(* IEC 61131-3 sources: daoli-st-library/DL_Base (part 14) *)

(* ---- FB_DL_MutexOwnerAudit.st ---- *)
(*
  FB_DL_MutexOwnerAudit  —  互斥锁所有权审计台账 / Mutex ownership audit ledger
  分类 Category : DL_Base
  码位 Code     : 16#01_0_02
  段位说明      : 01_0 段仅占 00/01（R38），02 起空穴，本件启用 02 格
  版本 Version  : 1.0.1
  来源 Source   : t0-8-sema — T0-8 行待挖子项「超时归还后的所有权审计」落地
  溯源 Origin   : clean-room 实现，未复制任何源码行
  功能 Function : 1) 只做「事后可追」审计出口，不改变加解锁语义：与 FB_DL_SemaMutex（互斥本体）
                  分工，本体管仲裁，本件管台账；
                  2) 记录持锁者标识 uOwnerCur、当前持有时长 fHoldCurSec、累计持有时长 uHoldTotalSec；
                  3) 计数台账：申请 / 正常释放 / 越权释放 / 超时强制归还四类，全部饱和计数不回绕；
                  4) 越权释放（无主时的释放沿）记故障级码并锁存，bReset 解除；
                  5) 超时强制归还由调用方把 FB_DL_SemaMutex.bTimedOut 单拍脉冲接入 bTimeoutForced。
  边界 Boundary : ① 本件不仲裁、不拒绝任何事件，只记录；仲裁语义全部由 FB_DL_SemaMutex 承载；
                  ② uDeltaTimeMs 为调用方注入的任务周期 [ms]，越界按上限钳位（防一次错误注入污染台账）；
                  R41 返修（R241）：饱和闸整体上移 UDINT 域——加法前预留量预检
                  （_uHoldMs / _uHoldTotMs 各自与 DL_MUA_MS_MAX - _uDtEff 比较），
                  判定值域 0..16#FFFF_F000 ms（约 49.7 天），以 10 ms 任务周期计约
                  4.29 亿拍可达，饱和分支真实可达，秒换算改纯 UDINT 整除，零降型路径；
                  ③ uOwnerIdClaim = 0 视为非法标识：照常记录持有但置信息级码 0302；
                  ④ 审计状态两相 CASE 全覆盖 + ELSE 兜底；无定时器/边沿以外的时序假设。
  依赖 Depends  : 仅 Standard.library（R_TRIG）；与 FB_DL_SemaMutex（已注册）仅状态语义对齐，不实例化
  码表 Error codes（本件格 01_0_02，子码步进 +0x100）:
    16#0001_0102 信息级：本拍记录到申请沿（持锁开始）
    16#0001_0202 故障级：越权释放（无主时的释放沿），锁存至 bReset
    16#0001_0302 信息级：申请者标识非法（uOwnerIdClaim = 0），记录照常完成
    16#0001_0402 信息级：超时强制归还事件已入账
    16#0001_0502 故障级：审计相位落 ELSE 兜底（非法相位 ID），强制回无主相并锁存

  修订历史 Revision :
    2026-11-19  v1.0.0  R39 首版（批次 1 · 序号 1）
    2026-11-19  v1.0.1  R40 5 抽终审挂账（不改逻辑）：⚠ 段 4 行 108 饱和闸「UDINT_TO_DINT(DL_MUA_SEC_MAX)」
                  对 16#FFFF_FFFE 做 DINT 降型溢出（回绕为负），乘积类型跨平台歧义；且 _uHoldTotMs
                  （UDINT ms）数学上不可能达到 SEC_MAX×1000 ms，秒级饱和分支永不按预期触发，返修轮处理。
    2026-11-19  v1.0.1  R41 P0-2 返修实施：删除「UDINT_TO_DINT(SEC_MAX) × 1000」降型比较与
                  不可达秒级闸，改为 UDINT 域加法前预留量预检（判定值域 0..16#FFFF_F000 ms，
                  可达性向量已写入边界②），秒换算改纯 UDINT 整除；新增常量 DL_MUA_MS_MAX，
                  DL_MUA_SEC_MAX 降级为文档口径不再参与比较。
*)

TYPE E_DL_MutexAuditState :
(
    eFree := 0,    // 无主：互斥空闲，等待申请沿 / Free, mutex idle, waiting for a claim edge
    eHeld := 10    // 有主：持锁审计中，累计持有时长 / Held, ownership held and hold time accumulating
);
END_TYPE

FUNCTION_BLOCK FB_DL_MutexOwnerAudit
VAR_INPUT
    bClaimEvt      : BOOL;                  // 申请事件沿（来自本体申请沿或其输入 CLK）[-] / Claim event edge from the mutex body
    bReleaseEvt    : BOOL;                  // 释放事件沿（来自本体释放沿或其输入 CLK）[-] / Release event edge from the mutex body
    bTimeoutForced : BOOL;                  // 超时强制归还脉冲，接 FB_DL_SemaMutex.bTimedOut 单拍输出 [-] / Forced timeout return pulse, wire SemaMutex.bTimedOut
    uOwnerIdClaim  : DINT := 0;             // 本次申请者标识 [ID]，0 = 非法（置信息码） / Claimer owner ID, 0 = illegal (info code)
    uDeltaTimeMs   : UDINT := 10;           // 任务周期注入 [ms]，越界按上限钳位 / Task cycle time injected by caller [ms]
    bReset         : BOOL := FALSE;         // 审计复位，上升沿清越权锁存（不清台账计数）/ Audit reset, rising edge clears the fault latch only
END_VAR
VAR_OUTPUT
    eState         : E_DL_MutexAuditState;  // 审计状态出口，段尾单点映射 / Audit state outlet
    bHeld          : BOOL;                  // 当前有主（与 eHeld 同源派生）/ Mutex currently held, derived from eHeld
    uOwnerCur      : DINT;                  // 当前持锁者标识 [ID]，无主时为 0 / Current owner ID, 0 when free
    fHoldCurSec    : REAL;                  // 当前连续持有时长 [s]，释放拍冻结到释放值 / Current continuous hold time [s], frozen at release
    uHoldTotalSec  : UDINT;                 // 累计持有时长 [s]，饱和不回绕 / Total accumulated hold time [s], saturating
    uClaimCnt      : UDINT;                 // 累计申请次数 [次]，饱和不回绕 / Total claim count [times], saturating
    uReleaseCnt    : UDINT;                 // 累计正常释放次数 [次]，饱和不回绕 / Total normal release count [times], saturating
    uUnauthRelCnt  : UDINT;                 // 累计越权释放次数 [次]，饱和不回绕 / Total unauthorized release count [times], saturating
    uTimeoutCnt    : UDINT;                 // 累计超时强制归还次数 [次]，饱和不回绕 / Total forced timeout return count [times], saturating
    uErrorId       : UDINT;                 // 事件码，0 = 无事件（故障级码锁存回放）/ Event code, 0 = none, fault codes latched and replayed
END_VAR
VAR
    rtClaim        : R_TRIG;                // 申请沿实例，主体首部无条件刷新 / Claim edge instance, refreshed unconditionally
    rtRelease      : R_TRIG;                // 释放沿实例，主体首部无条件刷新 / Release edge instance, refreshed unconditionally
    rtTimeout      : R_TRIG;                // 超时归还沿实例，主体首部无条件刷新 / Timeout edge instance, refreshed unconditionally
    rtReset        : R_TRIG;                // 复位沿实例，主体首部无条件刷新 / Reset edge instance, refreshed unconditionally
    _eState        : E_DL_MutexAuditState := E_DL_MutexAuditState.eFree;  // 内部审计相位（CASE 唯一写入目标）/ Internal audit phase, sole CASE target
    _uFault        : UDINT;                 // 故障码锁存寄存 / Latched fault code register
    _uInfo         : UDINT;                 // 本拍信息码，每拍重算 / Transient info code this cycle
    _uOwnerInt     : DINT := 0;             // 内部持锁者标识，对外经 uOwnerCur 镜像 / Internal owner register mirrored to uOwnerCur
    _uHoldMs       : UDINT := 0;            // 当前持有毫秒累加器 [ms] / Current hold millisecond accumulator
    _uHoldTotMs    : UDINT := 0;            // 累计持有毫秒累加器 [ms] / Total hold millisecond accumulator
    _uDtEff        : UDINT;                 // 钳位后的生效周期 [ms] / Clamped effective cycle time
END_VAR
VAR CONSTANT
    DL_MUA_DT_MAX     : UDINT := 60000;         // 单拍周期合理上限 [ms]，超出按上限入账 / Sane per-cycle cap [ms]
    DL_MUA_CNT_MAX    : UDINT := 16#FFFF_FFFE;  // 各计数饱和上限 [次]，加一永不回绕 / Counter saturation bound, increment never wraps
    DL_MUA_MS_PER_SEC : UDINT := 1000;          // 每秒毫秒数 [ms/s] / Milliseconds per second
    DL_MUA_SEC_MAX    : UDINT := 16#FFFF_FFFE;  // 秒级累计饱和上限 [s]，R41 起仅作文档口径，不再参与比较 / Second-level doc bound, not used in comparison since R41
    DL_MUA_MS_MAX     : UDINT := 16#FFFF_F000;  // 毫秒累加器饱和上限 [ms]，UDINT 域加法闸（约 49.7 天，10ms 周期约 4.29 亿拍可达）/ Millisecond accumulator saturation bound, UDINT-domain add gate
END_VAR

(* —— 段 0：边沿实例无条件周期刷新（R7 红线：严禁置于 IF/CASE 分支内） —— *)
rtClaim(CLK := bClaimEvt);                                        // 申请沿刷新，每拍必调
rtRelease(CLK := bReleaseEvt);                                    // 释放沿刷新，每拍必调
rtTimeout(CLK := bTimeoutForced);                                 // 超时归还沿刷新，每拍必调
rtReset(CLK := bReset);                                           // 复位沿刷新，每拍必调

(* —— 段 1：单拍量预清零（锁存量 _uFault 与台账计数不入清单，R187①） —— *)
_uInfo := 16#0000_0000;             // 信息码每拍重算
_uFault := _uFault;                 // 故障锁存码保持回放（禁同拍抹除，R187/R189）
uErrorId := 16#0000_0000;           // 事件码缺省无事件（段尾按锁存/信息单点回放）

(* —— 段 2：周期注入钳位（防御：一次错误注入不得污染台账） —— *)
IF uDeltaTimeMs > DL_MUA_DT_MAX THEN
    _uDtEff := DL_MUA_DT_MAX;       // 越界按上限钳位
ELSE
    _uDtEff := uDeltaTimeMs;        // 域内直通
END_IF

(* —— 段 3：复位沿（只清越权锁存，不清台账计数——台账是历史事实） —— *)
IF rtReset.Q THEN
    _uFault := 16#0000_0000;        // 清故障锁存码（唯一解除路径：bReset 上升沿）
END_IF

(* —— 段 4：持有时长累加（仅 eHeld 相累计；R41 P0-2 返修：饱和闸整体上移 UDINT 域，
     加法前预留量预检，判定值域 0..16#FFFF_F000 ms，无降型、无可达性缺口） —— *)
IF _eState = E_DL_MutexAuditState.eHeld THEN
    IF _uHoldMs <= DL_MUA_MS_MAX - _uDtEff THEN     // 加前预留量预检（当拍量判据，UDINT 域）
        _uHoldMs := _uHoldMs + _uDtEff;             // 当前持有累加 [ms]
    ELSE
        _uHoldMs := DL_MUA_MS_MAX;                  // 饱和钳位，永不回绕
    END_IF
    IF _uHoldTotMs <= DL_MUA_MS_MAX - _uDtEff THEN  // 同口径预检累计累加器（UDINT 域，零降型）
        _uHoldTotMs := _uHoldTotMs + _uDtEff;       // 累计持有累加 [ms]
    ELSE
        _uHoldTotMs := DL_MUA_MS_MAX;               // 累计饱和钳位，永不回绕
    END_IF
END_IF
fHoldCurSec := UDINT_TO_REAL(_uHoldMs) / UDINT_TO_REAL(DL_MUA_MS_PER_SEC);  // 当前持有换算秒（分母为常量恒非零）
uHoldTotalSec := _uHoldTotMs / DL_MUA_MS_PER_SEC;   // 累计秒整除换算（纯 UDINT 域，R241 零降型）

(* —— 段 5：审计相位机（只记录、不仲裁；出口在段 7） —— *)
CASE _eState OF

E_DL_MutexAuditState.eFree:
    IF rtRelease.Q THEN
        uUnauthRelCnt := uUnauthRelCnt + 1;     // 越权释放入账（无主时的释放沿）
        IF uUnauthRelCnt >= DL_MUA_CNT_MAX THEN
            uUnauthRelCnt := DL_MUA_CNT_MAX;    // 计数饱和防回绕
        END_IF
        _uFault := 16#0001_0202;                // 故障级：越权释放，锁存至 bReset
    ELSIF rtTimeout.Q THEN
        uTimeoutCnt := uTimeoutCnt + 1;         // 超时归还沿落在此相同样入账（本体已强制归还）
        IF uTimeoutCnt >= DL_MUA_CNT_MAX THEN
            uTimeoutCnt := DL_MUA_CNT_MAX;
        END_IF
        _uInfo := 16#0001_0402;                 // 信息级：超时归还已入账
    ELSIF rtClaim.Q THEN
        uClaimCnt := uClaimCnt + 1;             // 申请入账
        IF uClaimCnt >= DL_MUA_CNT_MAX THEN
            uClaimCnt := DL_MUA_CNT_MAX;
        END_IF
        IF uOwnerIdClaim = 0 THEN
            _uInfo := 16#0001_0302;             // 信息级：标识非法，记录照常
        ELSE
            _uInfo := 16#0001_0102;             // 信息级：持锁开始
        END_IF
        _uOwnerInt := uOwnerIdClaim;            // 记录持锁者标识（含非法 0，照实记录）
        _uHoldMs := 0;                          // 当前持有时长从零起算
        _eState := E_DL_MutexAuditState.eHeld;  // 进有主相
    END_IF

E_DL_MutexAuditState.eHeld:
    IF rtRelease.Q THEN
        uReleaseCnt := uReleaseCnt + 1;         // 正常释放入账
        IF uReleaseCnt >= DL_MUA_CNT_MAX THEN
            uReleaseCnt := DL_MUA_CNT_MAX;
        END_IF
        _uOwnerInt := 0;                        // 无主：标识清零
        _eState := E_DL_MutexAuditState.eFree;  // 回无主相（当前持有时长冻结在释放值）
    ELSIF rtTimeout.Q THEN
        uTimeoutCnt := uTimeoutCnt + 1;         // 超时强制归还有主相入账
        IF uTimeoutCnt >= DL_MUA_CNT_MAX THEN
            uTimeoutCnt := DL_MUA_CNT_MAX;
        END_IF
        _uInfo := 16#0001_0402;                 // 信息级：超时归还已入账
        _uOwnerInt := 0;                        // 强制归还：标识清零
        _eState := E_DL_MutexAuditState.eFree;  // 回无主相
    ELSIF rtClaim.Q THEN
        uClaimCnt := uClaimCnt + 1;             // 有主期间的申请沿照常入账（本体仲裁语义不变）
        IF uClaimCnt >= DL_MUA_CNT_MAX THEN
            uClaimCnt := DL_MUA_CNT_MAX;
        END_IF
    END_IF

ELSE
    _uFault := 16#0001_0502;                    // 故障级：非法相位 ID 兜底，锁存至 bReset
    _uOwnerInt := 0;                            // 无主侧强制清标识（安全侧）
    _eState := E_DL_MutexAuditState.eFree;      // 强制回无主相（自恢复，不锁死）

END_CASE

(* —— 段 6：派生输出每拍重写（名实同源） —— *)
bHeld := (_eState = E_DL_MutexAuditState.eHeld);            // 有主派生位
uOwnerCur := _uOwnerInt;                                     // 持锁者镜像输出

(* —— 段 7：事件码单点回放（故障锁存优先，信息码其次） —— *)
IF _uFault <> 16#0000_0000 THEN
    uErrorId := _uFault;            // 故障锁存码回放（不在故障态按当下输入重推）
ELSE
    uErrorId := _uInfo;             // 信息码
END_IF
eState := _eState;                  // 状态出口单点映射

END_FUNCTION_BLOCK

(* ---- FB_DL_OutputForcingBank.st ---- *)
(*==============================================================================
 * 组件名称 (Component)  : FB_DL_OutputForcingBank
 * 所属子库 (Sublibrary) : DL_Base
 * 当前版本 (Version)    : 1.0.0
 * 兼容性   (Platform)   : CODESYS 3.5+ / TwinCAT 3 / 汇川 InoProShop / 施耐德 Machine Expert
 *                         仅依赖 Standard.library（R_TRIG），零厂商私有库
 * 功能描述 (Function)   : 16 路输出强制库（调试/维修用）：每拍组合式裁决
 *                         abOut[i] = bAutoMode ∧ abForceSel[i] ? abForceVal[i]
 *                         : abAutoVal[i]；任一通道强制激活 → uForcingMask 位图
 *                         对应位置 1；强制撤除（abForceSel 下降沿）当拍无扰
 *                         回自动（组合式单拍重算，无斜坡无残留）；bAutoMode=
 *                         FALSE 时强制请求被拒（输出仍走自动值），拒收当拍置
 *                         信息码 eForceRej 并计数 uRejCnt。
 * 接口     (Interface)  : 输入 abAutoVal 16 路自动值、abForceSel 16 路强制选择、
 *                         abForceVal 16 路强制值、bAutoMode 自动模式许可；
 *                         输出 abOut 16 路裁决输出、uForcingMask 强制激活
 *                         位图（bit i=通道 i）、uRejCnt 强制拒收计数、
 *                         eErrCode 信息码、bError 故障标志（本件无故障级
 *                         条件，恒 FALSE，契约位保留）。
 * 边界     (Boundary)   : ① **属主边界（写死）：本件只做输出裁决，不接管安全
 *                         回路、不做强制权限管理**；安全回路强制归硬件层，
 *                         本件不得用于旁路安全联锁（头注释声明）。
 *                         ② 无扰回自动：撤除拍输出 = 自动值（组合式当拍生效，
 *                         无历史残留路径，规格指定）。
 *                         ③ 拒收计数用 R_TRIG 捕「拒收状态进入沿」计数（状态
 *                         电平不重复计数）；拒收期 uForcingMask 对应位保持 0
 *                         （强制未生效）。
 *                         ④ 通道定长 16（常量），FOR 界宽常量，无越界路径。
 *                         ⑤ R_TRIG 实例段 0 无条件周期调用（R6/R7）。
 *                         ⑥ 零全局耦合（无 GVL / VAR_EXTERNAL / 物理地址）。
 * 分工声明 (Scope)      : 与 `FB_DL_OverrideSelector` 分工：模拟量超驰选择归
 *                         那件、数字量强制库归本件；与 `FB_DL_InterlockMatrix`
 *                         分工：联锁矩阵归那件（安全语义），本件为非安全
 *                         调试设施。
 * 来源标签 (Source Tag) : 自研线（输出强制裁决为道莅防御性实现）
 * 码表     (Codes)      : 本件不占用任何全局数字码位。出口为 BOOL 数组 +
 *                         WORD 位图 + UDINT 计数 + ENUM 信息码；数字码位待
 *                         主控收口阶段统一派号。
 * 红线自检 (Redline)    : R1 ✓ 零 GVL/VAR_EXTERNAL ｜ R2 ✓ 零 %I/%Q/%M ｜ R3 ✓ 纯 IEC 61131-3
 *                         R4 ✓ 拒收沿计数 + 无扰回自动 + 位图单源 ｜ R5 ✓ 声明逐行同行双语注释
 *                         R6 N/A（无 ENUM 状态机） ｜ R7 ✓ 一 R_TRIG 段 0 无条件刷新
 * 修订历史 (Revision)   : 2026-11-20  v1.0.0  R50 首版（批次 3 · 序号 12）
 * 验收向量 (Acceptance) : ① bAutoMode=TRUE，abForceSel[3]=TRUE，abForceVal[3]=
 *                         TRUE，abAutoVal[3]=FALSE → abOut[3]=TRUE，
 *                         uForcingMask.bit3=1；② abForceSel[3] 撤除当拍：
 *                         abOut[3]=abAutoVal[3]=FALSE（无扰回自动），bit3=0；
 *                         ③ bAutoMode=FALSE 且 abForceSel[5] 置位 → abOut[5]
 *                         =abAutoVal[5]（强制被拒），uRejCnt+1，
 *                         eErrCode=eForceRej。
 *==============================================================================*)

(*-----------------------------------------------------------------------------
 * 枚举: E_DL_OfbErr（信息码；拒收走信息级，不置 bError）
 *----------------------------------------------------------------------------*)
TYPE E_DL_OfbErr :
(
    eOk       := 0,   // 无拒收 / No rejection
    eForceRej := 1    // 信息级：存在被拒强制通道（bAutoMode=FALSE，见 uRejCnt） / Info: forced channels rejected
);
END_TYPE

FUNCTION_BLOCK FB_DL_OutputForcingBank
VAR_INPUT
    abAutoVal  : ARRAY[0..15] OF BOOL;   // 16 路自动值（正常输出源） [-] / Sixteen auto values
    abForceSel : ARRAY[0..15] OF BOOL;   // 16 路强制选择 [-] / Sixteen force selects
    abForceVal : ARRAY[0..15] OF BOOL;   // 16 路强制值 [-] / Sixteen force values
    bAutoMode  : BOOL := TRUE;           // 自动模式许可（FALSE=强制被拒） [-] / Auto-mode permission
END_VAR
VAR_OUTPUT
    abOut        : ARRAY[0..15] OF BOOL; // 16 路裁决输出 [-] / Sixteen arbitrated outputs
    uForcingMask : WORD;                 // 强制激活位图（bit i=通道 i 强制生效） [-] / Forcing bitmap
    uRejCnt      : UDINT := 0;           // 强制拒收进入沿计数（防回绕） [次] / Rejection entry count
    eErrCode     : E_DL_OfbErr;          // 信息码出口 / Info code outlet
    bError       : BOOL;                 // 故障标志（本件恒 FALSE，契约位） [-] / Error flag, contract pin, always FALSE
END_VAR
VAR
    _uMask    : WORD;                    // 位图内部单源（与出口同源） / Bitmap internal source
    _bAnyRej  : BOOL;                    // 存在拒收通道当拍量 [-] / Any rejected channel
    i         : DINT;                    // 通道循环索引 / Channel loop index
    rtRej     : R_TRIG;                  // 拒收进入沿实例，段 0 无条件调用 / Rejection entry edge instance
END_VAR
VAR CONSTANT
    DL_OFB_NMAX : DINT := 16;            // 通道定长 [路] / Fixed channel count
    DL_OFB_BIT0 : WORD := 1;             // bit0 基准掩码 [-] / Bit zero base mask
    DL_OFB_UDMAX: UDINT := 4294967295;   // 拒收计数饱和点（防回绕） [次] / Rejection counter ceiling
END_VAR

(* —— 段 0：拒收沿实例无条件周期刷新（R6/R7） —— *)
rtRej(CLK := (NOT bAutoMode) AND (abForceSel[0] OR abForceSel[1] OR abForceSel[2]
       OR abForceSel[3] OR abForceSel[4] OR abForceSel[5] OR abForceSel[6]
       OR abForceSel[7] OR abForceSel[8] OR abForceSel[9] OR abForceSel[10]
       OR abForceSel[11] OR abForceSel[12] OR abForceSel[13] OR abForceSel[14]
       OR abForceSel[15]));              // 拒收进入沿（任一强制选择 ∧ 非自动模式），每拍必调 / Rejection entry edge, every scan

(* —— 段 1：拒收沿计数（防回绕） —— *)
IF rtRej.Q THEN
    IF uRejCnt < DL_OFB_UDMAX THEN
        uRejCnt := uRejCnt + 1;          // 拒收进入沿计数 / Count rejection entry
    END_IF
END_IF

(* —— 段 2：16 路组合式裁决（强制生效闸：bAutoMode ∧ abForceSel；撤除当拍无扰回自动） —— *)
_uMask := 0;                             // 位图当拍重建（单源） / Rebuild bitmap per scan
_bAnyRej := FALSE;                       // 拒收量预清 / Rejection preset
FOR i := 0 TO (DL_OFB_NMAX - 1) DO
    IF bAutoMode AND abForceSel[i] THEN
        abOut[i] := abForceVal[i];       // 强制生效：输出强制值 / Forced: force value
        _uMask := _uMask OR SHL(DL_OFB_BIT0, i);   // 记激活位（i∈[0,15] 位宽内） / Set forcing bit
    ELSE
        abOut[i] := abAutoVal[i];        // 自动值直通（含强制撤除当拍与拒收通道） / Auto pass-through
        IF abForceSel[i] THEN
            _bAnyRej := TRUE;            // 强制请求被拒（bAutoMode=FALSE） / Force rejected
        END_IF
    END_IF
END_FOR

(* —— 段 3：出口单点映射（名实双出口同源，R191） —— *)
uForcingMask := _uMask;                  // 位图出口 / Bitmap outlet
IF _bAnyRej THEN
    eErrCode := E_DL_OfbErr.eForceRej;   // 信息级（不置 bError） / Info code
ELSE
    eErrCode := E_DL_OfbErr.eOk;         // 正常 / Normal
END_IF
bError := FALSE;                         // 本件无故障级条件（头注释声明） / No fault-level condition

END_FUNCTION_BLOCK

(* ---- FB_DL_ParamSnapshotRestore.st ---- *)
// FB_DL_ParamSnapshotRestore v1.0.0
// 开源溯源：self-cleanroom / 参数管理族
(*
  道莅工业代码库 | DL_Base | FB_DL_ParamSnapshotRestore
  版本: 1.0.0 | 日期: 2026-11-23 | 轮次: R75
  功能: 参数快照/一键回滚：双缓冲（快照写入非活动缓冲区并切换），回滚时
        把最近有效快照整组复制回输出组；快照序号累加供追溯
  邻件关系: 与 DeviceParamVerify / DeviceParamWrite（参数校验/写入）同族 ——
            差异点：校验/写入件为单参数级在线动作，本件为整组快照与
            历史回滚（双缓冲），互不重叠
  时序契约: bSnap 上升沿写快照（双缓冲切换）；bRestore 上升沿回滚最近快照；
            两沿同拍时快照优先（先存后回滚，本拍回滚的是新快照）
*)
FUNCTION_BLOCK FB_DL_ParamSnapshotRestore
VAR_INPUT
    bSnap      : BOOL := FALSE;              // 快照触发（上升沿）/ Snapshot trigger, rising edge
    bRestore   : BOOL := FALSE;              // 回滚触发（上升沿）/ Restore trigger, rising edge
    aParamIn   : ARRAY[1..16] OF REAL;       // 参数输入组 [工程单位] / Parameter input group
    nCount     : INT := 16;                  // 有效参数个数 [个]，域 1..16 / Valid parameter count
END_VAR
VAR_OUTPUT
    aParamOut  : ARRAY[1..16] OF REAL;       // 参数输出组（回滚目标）[工程单位] / Parameter output group, restore target
    nSnapSeq   : UDINT;                      // 快照序号（每次快照 +1）/ Snapshot sequence number
    bSnapDone  : BOOL;                       // 快照完成脉冲（单拍自清）/ Snapshot done pulse, one cycle
    bRestDone  : BOOL;                       // 回滚完成脉冲（单拍自清）/ Restore done pulse, one cycle
    bHasSnap   : BOOL;                       // 存在可用快照 [-] / Valid snapshot available
    bValid     : BOOL;                       // 组态有效回执 [-] / Config validity receipt
    bError     : BOOL;                       // 故障标志（计数非法）/ Fault flag (invalid count)
    uErrorId   : UDINT;                      // 事件码，0 = 无事件；16#0002_2101 = 计数非法 / Event code
END_VAR
VAR
    rtrSnap    : R_TRIG;                     // 快照沿检测（每拍无条件刷新）/ Snapshot edge, refreshed every cycle
    rtrRest    : R_TRIG;                     // 回滚沿检测（每拍无条件刷新）/ Restore edge, refreshed every cycle
    aBufA      : ARRAY[1..16] OF REAL;       // 缓冲区 A [工程单位] / Buffer A
    aBufB      : ARRAY[1..16] OF REAL;       // 缓冲区 B [工程单位] / Buffer B
    bActiveA   : BOOL;                       // 最近快照在缓冲区 A [-] / Latest snapshot in buffer A
    i          : INT;                        // 复制循环索引 [个] / Copy loop index
    nCnt       : INT;                        // 钳位后生效个数 [个] / Effective clamped count
END_VAR

// —— 段 0：实例无条件刷新 + 输出缺省 —— //
rtrSnap(CLK := bSnap);                       // 快照沿每拍刷新 / Snapshot edge refreshed
rtrRest(CLK := bRestore);                    // 回滚沿每拍刷新 / Restore edge refreshed
bSnapDone := FALSE;                          // 快照脉冲单拍自清 / Snapshot pulse self-clearing
bRestDone := FALSE;                          // 回滚脉冲单拍自清 / Restore pulse self-clearing

// —— 段 1：计数域闸（下标判界，R4） —— //
bValid := (nCount >= 1) AND (nCount <= 16);  // 计数域 1..16 / Count domain
IF NOT bValid THEN
    bError   := TRUE;                        // 故障级：计数非法 / Fault level: illegal count
    uErrorId := 16#0002_2101;                // 故障码（21xx 步进）/ Fault code
    RETURN;                                  // 非法计数不动作 / No action on illegal count
END_IF
bError   := FALSE;                           // 组态恢复：故障清零（解除路径）/ Fault cleared
uErrorId := 16#0000;                         // 事件码清零 / Event code cleared
nCnt := nCount;                              // 生效个数 / Effective count

// —— 段 2：快照沿（双缓冲：写入非活动区并切换；同拍快照优先于回滚） —— //
IF rtrSnap.Q THEN
    IF bActiveA THEN                         // 当前最近快照在 A：写入 B / Latest in A: write to B
        FOR i := 1 TO nCnt DO                 // 逐元素复制（i ≤ nCnt ≤ 16 判界安全）/ Copy elements, index safe
            aBufB[i] := aParamIn[i];
        END_FOR
        bActiveA := FALSE;                   // 最近快照切到 B / Latest now in B
    ELSE                                     // 当前最近快照在 B：写入 A / Latest in B: write to A
        FOR i := 1 TO nCnt DO
            aBufA[i] := aParamIn[i];
        END_FOR
        bActiveA := TRUE;                    // 最近快照切到 A / Latest now in A
    END_IF
    bHasSnap := TRUE;                        // 存在可用快照 / Snapshot available
    nSnapSeq := nSnapSeq + 1;                // 快照序号累加（UDINT 回绕无害）/ Sequence increments
    bSnapDone := TRUE;                       // 快照完成脉冲 / Snapshot done pulse
END_IF

// —— 段 3：回滚沿（复制最近快照到输出组） —— //
IF rtrRest.Q AND bHasSnap THEN               // 有快照才回滚 / Restore only with snapshot
    IF bActiveA THEN                         // 最近快照在 A / Latest in A
        FOR i := 1 TO nCnt DO
            aParamOut[i] := aBufA[i];
        END_FOR
    ELSE                                     // 最近快照在 B / Latest in B
        FOR i := 1 TO nCnt DO
            aParamOut[i] := aBufB[i];
        END_FOR
    END_IF
    bRestDone := TRUE;                       // 回滚完成脉冲 / Restore done pulse
END_IF
END_FUNCTION_BLOCK

(* ---- FB_DL_PrbsSignal.st ---- *)
(*
  Name        : FB_DL_PrbsSignal
  Category    : DL_Base
  Version     : 1.0.0
  Purpose     : PRBS 伪随机二进序列激励发生（LFSR 整数实现，阶数 4..31 抽头表），供回路辨识/继电器整定的持续激励源；/ PRBS pseudo-random binary sequence excitation generator (integer LFSR, degree 4..31 tap table) for loop identification and relay tuning
  溯源        : 借 oscat-basic 的 PRBS 行为定义组织，clean-room 实现
  Boundary    : ① 抽头多项式合法域校验：阶数 4..31 之外的阶数锁存故障（抽头表 CASE 全覆盖 + ELSE 兜底）；
                ② LFSR 全零态检测：每步推进前遇全零强制注入 1（防死序列）；
                ③ 使能撤除保持相位与序列值，重使能不重启序列；仅 bRestart 上升沿显式重载种子重启；
                ④ 输出脉冲宽度以扫描周期为时基（每 nBitScan 拍推进一位），nBitScan 钳位下限 ≥ 2；
                ⑤ 种子 0 视为非法（与全零态同源），组态期锁存故障；
                ⑥ 零外部全局、零物理地址，纯整数实现跨平台移植。
*)
TYPE E_DL_PbsState :
(
    eIdle  := 0,                             (* 未使能（相位保持） / Disabled, phase held *)
    eRun   := 10,                            (* 序列激励运行 / Sequence running *)
    eFault := 90                             (* 故障锁存相 / Fault latched *)
);
END_TYPE

TYPE E_DL_PbsCause :
(
    eNone      := 0,                         (* 无故障成因 / No cause *)
    eCfgIllegal:= 1,                        (* 组态非法：阶数/种子/位宽越域 / Illegal config *)
    ePhaseBad  := 2                         (* 非法相位兜底 / Illegal phase fallback *)
);
END_TYPE

FUNCTION_BLOCK FB_DL_PrbsSignal
VAR_INPUT
    nDegree : INT := 31;                     (* LFSR 阶数，域 4..31 [阶] / LFSR degree *)
    nSeed   : DWORD := DWORD#16#ACE1;        (* 种子（0 非法）[-] / Seed, zero illegal *)
    nBitScan: INT := 10;                     (* 每位驻留扫描拍数，域 >= 2 [拍] / Bit dwell in scans *)
    bEnable : BOOL := TRUE;                  (* 使能（撤除保持相位）[-] / Enable, phase held on disable *)
    bRestart: BOOL := FALSE;                 (* 重启命令，上升沿重载种子 [-] / Restart command, edge reload seed *)
    bReset  : BOOL := FALSE;                 (* 复位命令，上升沿清故障与序列 [-] / Reset command *)
END_VAR
VAR_OUTPUT
    bOut    : BOOL;                          (* PRBS 位输出（当前 LFSR 最低位）[-] / PRBS bit output *)
    nBitCnt : UDINT;                         (* 已推进位数（饱和，诊断）[位] / Bits advanced, saturated *)
    eState  : E_DL_PbsState;                 (* 状态出口 / State outlet *)
    eCause  : E_DL_PbsCause;                 (* 故障成因出口（R190 归因唯一） / Fault cause outlet *)
    bError  : BOOL;                          (* 故障锁存标志 [-] / Fault latch flag *)
END_VAR
VAR
    _eState : E_DL_PbsState := E_DL_PbsState.eIdle;  (* 内部相位（CASE 唯一写入目标） / Internal phase *)
    _eCause : E_DL_PbsCause := E_DL_PbsCause.eNone;  (* 故障成因锁存量 / Latched cause *)
    rtReset : R_TRIG;                        (* 复位沿实例，段 0 无条件调用 / Reset edge instance *)
    rtRestart: R_TRIG;                       (* 重启沿实例，段 0 无条件调用 / Restart edge instance *)
    _bFault : BOOL;                          (* 故障锁存位 / Latched fault bit *)
    _bCfgBad: BOOL;                          (* 组态非法当拍量 / Illegal config this scan *)
    _nLfsr  : DWORD;                         (* LFSR 状态寄存器（整数实现）[-] / LFSR state register *)
    _nDegree: INT := 1;                      (* 当前反馈阶次（1 起，用于 SHL 位序）[-] / Current feedback degree, 1-based shift index *)
    _nTapMsk: DWORD;                         (* 抽头掩码（CASE 表派生）[-] / Tap mask from table *)
    _bFb    : BOOL;                          (* 反馈位异或累加量 [-] / Feedback parity *)
    _bZero  : BOOL;                          (* 全零态检测当拍量 / All-zero state detect *)
    _nDiv   : INT;                           (* 扫描分频计数器 [拍] / Scan divider counter *)
    _nDwell : INT;                           (* 钳位后生效位驻留拍数 [拍] / Clamped bit dwell *)
    _i      : INT;                           (* 抽头位扫描游标 [位] / Tap bit cursor *)
END_VAR
VAR CONSTANT
    DL_PBS_NMIN : INT   := 4;                (* 阶数下限（边界①）[阶] / Degree lower bound *)
    DL_PBS_NMAX : INT   := 31;               (* 阶数上限（边界①）[阶] / Degree upper bound *)
    DL_PBS_DMIN : INT   := 2;                (* 位驻留下限（边界④）[拍] / Dwell lower bound *)
    DL_PBS_CNTMAX: UDINT := 4294967295;      (* 推进计数饱和上限（R28）[位] / Count saturation cap *)
    DL_PBS_ONE  : DWORD := DWORD#1;          (* 位掩码常量 1 [-] / Bit mask one *)
END_VAR

(* —— 段 0：当拍判据派生 + 实例无条件刷新（R228A） —— *)
_bCfgBad := (nDegree < DL_PBS_NMIN) OR (nDegree > DL_PBS_NMAX)          (* 阶数域闸（边界①） / Degree gate *)
            OR (nSeed = DWORD#0)                                        (* 种子零非法闸（边界⑤） / Seed gate *)
            OR (nBitScan < DL_PBS_DMIN);                                (* 位驻留下限闸（边界④） / Dwell gate *)
rtReset(CLK := bReset);                                  (* 复位沿每拍必调 / Reset edge every scan *)
rtRestart(CLK := bRestart);                              (* 重启沿每拍必调 / Restart edge every scan *)
_nDwell := nBitScan;                                     (* 驻留拍数初值 / Dwell init *)
IF _nDwell < DL_PBS_DMIN THEN
    _nDwell := DL_PBS_DMIN;                              (* 驻留钳位下限（防 0 拍高频抖动） / Dwell clamp *)
END_IF

(* —— 段 0B：抽头掩码 CASE 表（本原多项式，位号 = 抽头位 - 1；每拍派生，全枚举覆盖 + ELSE 兜底，红线 5/6） —— *)
CASE nDegree OF
    4 : _nTapMsk := DWORD#16#0000000C;                   (* 抽头 4,3 → 位 3,2 / Taps 4,3 *)
    5 : _nTapMsk := DWORD#16#00000014;                   (* 抽头 5,3 → 位 4,2 / Taps 5,3 *)
    6 : _nTapMsk := DWORD#16#00000030;                   (* 抽头 6,5 → 位 5,4 / Taps 6,5 *)
    7 : _nTapMsk := DWORD#16#00000060;                   (* 抽头 7,6 → 位 6,5 / Taps 7,6 *)
    8 : _nTapMsk := DWORD#16#000000B8;                   (* 抽头 8,6,5,4 → 位 7,5,4,3 / Taps 8,6,5,4 *)
    9 : _nTapMsk := DWORD#16#00000110;                   (* 抽头 9,5 → 位 8,4 / Taps 9,5 *)
    10: _nTapMsk := DWORD#16#00000240;                   (* 抽头 10,7 → 位 9,6 / Taps 10,7 *)
    11: _nTapMsk := DWORD#16#00000500;                   (* 抽头 11,9 → 位 10,8 / Taps 11,9 *)
    12: _nTapMsk := DWORD#16#00000820;                   (* 抽头 12,6 → 位 11,5 / Taps 12,6 *)
    13: _nTapMsk := DWORD#16#0000100D;                   (* 抽头 13,4,3,1 → 位 12,3,2,0 / Taps 13,4,3,1 *)
    14: _nTapMsk := DWORD#16#00002015;                   (* 抽头 14,5,3,1 → 位 13,4,2,0 / Taps 14,5,3,1 *)
    15: _nTapMsk := DWORD#16#00006000;                   (* 抽头 15,14 → 位 14,13 / Taps 15,14 *)
    16: _nTapMsk := DWORD#16#0000B400;                   (* 抽头 16,14,13,11 → 位 15,13,12,10 / Taps 16,14,13,11 *)
    17: _nTapMsk := DWORD#16#00012000;                   (* 抽头 17,14 → 位 16,13 / Taps 17,14 *)
    18: _nTapMsk := DWORD#16#00020400;                   (* 抽头 18,11 → 位 17,10 / Taps 18,11 *)
    19: _nTapMsk := DWORD#16#00040023;                   (* 抽头 19,6,2,1 → 位 18,5,1,0 / Taps 19,6,2,1 *)
    20: _nTapMsk := DWORD#16#00090000;                   (* 抽头 20,17 → 位 19,16 / Taps 20,17 *)
    21: _nTapMsk := DWORD#16#00140000;                   (* 抽头 21,19 → 位 20,18 / Taps 21,19 *)
    22: _nTapMsk := DWORD#16#00300000;                   (* 抽头 22,21 → 位 21,20 / Taps 22,21 *)
    23: _nTapMsk := DWORD#16#00420000;                   (* 抽头 23,18 → 位 22,17 / Taps 23,18 *)
    24: _nTapMsk := DWORD#16#00E10000;                   (* 抽头 24,23,22,17 → 位 23,22,21,16 / Taps 24,23,22,17 *)
    25: _nTapMsk := DWORD#16#01200000;                   (* 抽头 25,22 → 位 24,21 / Taps 25,22 *)
    26: _nTapMsk := DWORD#16#2000023;                    (* 抽头 26,6,2,1 → 位 25,5,1,0 / Taps 26,6,2,1 *)
    27: _nTapMsk := DWORD#16#4000013;                    (* 抽头 27,5,2,1 → 位 26,4,1,0 / Taps 27,5,2,1 *)
    28: _nTapMsk := DWORD#16#09000000;                   (* 抽头 28,25 → 位 27,24 / Taps 28,25 *)
    29: _nTapMsk := DWORD#16#14000000;                   (* 抽头 29,27 → 位 28,26 / Taps 29,27 *)
    30: _nTapMsk := DWORD#16#30000000;                   (* 抽头 30,29 → 位 29,28 / Taps 30,29 *)
    31: _nTapMsk := DWORD#16#48000000;                   (* 抽头 31,28 → 位 30,27 / Taps 31,28 *)
    ELSE
        _nTapMsk := DWORD#0;                             (* 越域阶数：掩码清零（域闸已另行锁故障） / Out-of-domain degree *)
END_CASE

(* —— 段 1：单拍量预清零（R107） —— *)
bOut := FALSE;                                           (* 位输出预清（派生拍覆盖） / Bit output preset *)
_bFb := FALSE;                                           (* 反馈奇偶累加清零 / Feedback parity clear *)
_bZero := FALSE;                                         (* 全零态检测清零 / Zero detect clear *)

(* —— 段 2：复位沿处理（作用域：清故障 + 清序列状态 + 迁 eIdle，R283 逐项声明） —— *)
IF rtReset.Q THEN
    _bFault := FALSE;                                    (* 清故障锁存 / Clear fault *)
    _eCause := E_DL_PbsCause.eNone;                      (* 清成因 / Clear cause *)
    _nLfsr := DWORD#0;                                   (* 清序列寄存器 / Clear LFSR register *)
    _nDiv := 0;                                          (* 清分频计数 / Clear divider *)
    nBitCnt := UDINT#0;                                  (* 清推进计数出口 / Clear bit count *)
    bOut := FALSE;                                       (* 清位输出出口 / Clear bit output *)
    _eState := E_DL_PbsState.eIdle;                      (* 迁未使能相 / Back to idle *)
END_IF

(* —— 段 3：组态故障锁存（锁存至复位沿，R189） —— *)
IF _bCfgBad AND NOT _bFault THEN
    _bFault := TRUE;                                     (* 锁存故障位 / Latch fault *)
    _eCause := E_DL_PbsCause.eCfgIllegal;                (* 成因：组态非法 / Cause illegal config *)
    _eState := E_DL_PbsState.eFault;                     (* 同步迁故障相 / Migrate to fault *)
END_IF

(* —— 段 4：CASE 主状态机（ELSE 兜底迁 eFault，红线 6） —— *)
CASE _eState OF
    E_DL_PbsState.eIdle:                                 (* 未使能：相位与序列值保持（边界③） / Disabled, phase held *)
        bOut := FALSE;                                   (* 失能位输出确定值 0 / Disabled bit output zero *)
        _nDiv := 0;                                      (* 失能清分频计数（重使能重新计时） / Clear divider *)
        IF bEnable AND NOT _bFault THEN
            _nLfsr := nSeed;                             (* 使能迁入拍装载种子（相位起点） / Load seed at entry *)
            _nDiv := 0;                                  (* 分频计数归零 / Divider zero *)
            _eState := E_DL_PbsState.eRun;               (* 进入运行相 / Enter running *)
        END_IF
    E_DL_PbsState.eRun:                                  (* 运行相：分频推进 + 抽头反馈 / Running *)
        IF NOT bEnable THEN
            _eState := E_DL_PbsState.eIdle;              (* 失能回未使能（相位保持不重启） / Back to idle *)
        ELSE
            IF rtRestart.Q THEN
                _nLfsr := nSeed;                         (* 显式重启重载种子（边界③） / Explicit restart reload *)
                _nDiv := 0;                              (* 分频计数归零 / Divider zero *)
            END_IF
            _nDiv := _nDiv + 1;                          (* 分频计数递进 / Divider advance *)
            IF _nDiv >= _nDwell THEN                     (* 满驻留拍数推进一位（边界④） / Advance one bit *)
                _nDiv := 0;                              (* 分频计数回零 / Divider reset *)
                IF _nLfsr = DWORD#0 THEN
                    _bZero := TRUE;                      (* 全零态检测（边界②） / All-zero detect *)
                END_IF
                IF _bZero THEN
                    _nLfsr := DL_PBS_ONE;                (* 全零强制注入 1 防死序列（边界②） / Inject one on zero *)
                END_IF
                _bFb := FALSE;                           (* 反馈奇偶清零重算 / Parity clear recompute *)
                FOR _i := 0 TO 30 DO                     (* 抽头位扫描（0..30 有界） / Tap bit scan *)
                    IF (_nTapMsk AND SHL(DL_PBS_ONE, _i)) <> DWORD#0 THEN    (* 该位在抽头集内 / Bit in tap set *)
                        IF (_nLfsr AND SHL(DL_PBS_ONE, _i)) <> DWORD#0 THEN  (* 该位为 1 / Bit is one *)
                            _bFb := NOT _bFb;            (* 异或奇偶累加 / XOR parity accumulate *)
                        END_IF
                    END_IF
                END_FOR
                _nLfsr := SHR(_nLfsr, 1);                (* 右移推进 / Shift advance *)
                IF _bFb THEN
                    _nLfsr := _nLfsr OR SHL(DL_PBS_ONE, _nDegree - 1);   (* 反馈位插入最高位 / Insert feedback bit *)
                END_IF
                IF nBitCnt < DL_PBS_CNTMAX THEN
                    nBitCnt := nBitCnt + UDINT#1;        (* 推进计数净额累加（饱和） / Bit count accumulate *)
                END_IF
            END_IF
            bOut := (_nLfsr AND DL_PBS_ONE) = DL_PBS_ONE;    (* 位输出 = LFSR 最低位（位等比较） / Output = LFSR LSB *)
        END_IF
    E_DL_PbsState.eFault:                                (* 故障相：冻结保持，仅复位沿出 / Fault *)
        ;                                                (* 锁存回放（R28） / Replay from latch *)
    ELSE                                                 (* 非法相位兜底迁安全态 / Illegal phase fallback *)
        _eState := E_DL_PbsState.eFault;                 (* 迁故障相 / To fault *)
        _bFault := TRUE;                                 (* 同步锁存 / Latch *)
        _eCause := E_DL_PbsCause.ePhaseBad;              (* 成因：非法相位 / Cause illegal phase *)
END_CASE

(* —— 段 5：出口映射（bError/eState 同源，R191） —— *)
bError := _bFault;                                       (* 故障标志镜像 / Fault flag mirror *)
eState := _eState;                                       (* 状态出口 / State outlet *)
eCause := _eCause;                                       (* 成因出口 / Cause outlet *)
END_FUNCTION_BLOCK

(* ---- FB_DL_PulseGenerator.st ---- *)
(*==============================================================================
 * 组件名称 (Component)  : FB_DL_PulseGenerator
 * 所属子库 (Sublibrary) : DL_Base
 * 当前版本 (Version)    : 1.0.1
 * 兼容性   (Platform)   : CODESYS 3.5 / TwinCAT 3 / 汇川 InoProShop / Machine Expert
 *                         仅依赖 Standard.library（TON / R_TRIG），时间-实数换算用
 *                         IEC 标准 TIME_TO_REAL / REAL_TO_TIME 转换族（毫秒语义）
 * 功能描述 (Function)   : 周期与占空比运行时可调的方波发生器，支持相位复位与禁用重启。
 *                         用 ENUM 相位状态机（高相位 / 低相位）+ 单个 TON 实现，
 *                         不引入任何平台时刻函数，行为与扫描周期严格耦合、可预期。
 *                         占空比 0 与 1 分别退化为恒低与恒高（显式分支输出，不靠相位机碰运气）；
 *                         周期设下限防止脉冲窄到下游边沿检测丢沿；
 *                         越界参数钳位后继续运行并告警，绝不停机。
 * 开源溯源 (Origin)     : 原创实现。方波 / 占空比调制为公开经典需求；
 *                         本库刻意放弃"记录时刻再比较"的实现路线，
 *                         改用标准定时器 + 相位状态机，未复制任何源码。
 * 本文件内含       : TYPE  E_DL_PulsePhase（配套枚举，归属 DL_Base）
 *                    FB    FB_DL_PulseGenerator
 * 依赖     (Depends)    : 无 DL_ 内部依赖；Standard.library: TON / R_TRIG
 * 红线自检 (Redline)    : R1 ✓ 禁用全局存储与物理寻址 ｜ R2 ✓ 无地址直写
 *                         R3 ✓ 纯 IEC 61131-3（时间换算走标准转换族）｜ R4 ✓ 容差判等 + 周期钳位 + 进度钳位
 *                         R5 ✓ 全变量中英双语同行注释 ｜ R6 ✓ 四态 ENUM + CASE + ELSE 兜底
 *                         R7 ✓ 两实例主体最前部无条件刷新 ｜ R8 ✓ 上下限与容差全常量化
 *
 * 【周期下限的存在理由 / Why the lower period bound exists（边界 B3）】
 *   脉宽低于两个任务周期时，下游边沿检测在扫描采样的离散化下必然丢沿，
 *   表现为"下游偶尔少计一次"。故下限设为 2ms，低于下限一律钳位并告警。
 *
 * 【平台收窄预案 / Platform narrowing contingency（边界 B5，R11）】
 *   时间-实数换算使用 IEC 标准转换族；若目标平台实测不支持该转换族，
 *   按规格书 P4 预案收窄：删去 fProgress 引脚并以整型毫秒中间量实现时长拆分，
 *   届时须在头注释追加收窄依据与影响说明。当前版本未启用收窄。
 *
 * 修订历史 (Revision)   :
 *   2026-11-14  v1.0.0  首版入库（Phase 1 第二轮 · Level 0 批次 B）
 *   2026-11-14  v1.0.1  修复换相后相位定时器不清零缺陷：标准定时器仅在本体输入为
 *                       FALSE 时清已计时，换相时只改预设值不会清零，低相位带着
 *                       高相位残值起算——占空比 0.5 时低相位塌缩为一个扫描周期，
 *                       占空比 0.3 时周期由 1000ms 变成 700ms。改为换相后追加一拍
 *                       断开输入（断拍屏蔽标志延后一拍提交），相位时长恢复设计值。
 *============================================================================*)

(*-----------------------------------------------------------------------------
 * 枚举: E_DL_PulsePhase（归属 DL_Base，与 FB_DL_PulseGenerator 同文件）
 * 含义: 方波相位状态。数值步长留空位便于后续插态而不破坏已有工程。
 *----------------------------------------------------------------------------*)
TYPE E_DL_PulsePhase :
(
    eInit  := 0,     // 上电/未使能首态：输出低，等待使能 / Power-up or disabled, output low and waits for enable
    eHigh  := 10,    // 高电平相位：持续 tHighTime / High phase lasting tHighTime
    eLow   := 20,    // 低电平相位：持续 tLowTime / Low phase lasting tLowTime
    eFault := 99     // 故障锁定：输出强制低 / Fault latched, output forced low
);
END_TYPE

FUNCTION_BLOCK FB_DL_PulseGenerator
VAR_INPUT
    bEnable     : BOOL := TRUE;       // 使能，FALSE 时输出 FALSE 并复位相位 / Enable, FALSE forces the output low and resets the phase
    tPeriod     : TIME := T#1S;       // 周期 [ms]，合法域为下限至上限 / Period [ms], valid range between the bounds
    fDutyCycle  : REAL := 0.5;        // 占空比 [0..1]，0 = 恒低，1 = 恒高 / Duty ratio [0..1], 0 = always low, 1 = always high
    bPhaseReset : BOOL;               // 上升沿：相位回高电平起点 / Rising edge: restart at the high phase
END_VAR
VAR_OUTPUT
    bPulseOut   : BOOL;     // 方波输出 / Square-wave output
    fProgress   : REAL;     // 当前周期进度 [0..1] / Cycle progress [0..1]
    bError      : BOOL;     // 故障/告警标志 / Fault or warning flag
    uErrorId    : UDINT;    // 故障码，0 = 无故障 / Error code, 0 = no error
END_VAR
VAR
    fbTonPhase  : TON;                // 相位计时器 / Phase timer
    fbTrigReset : R_TRIG;             // 相位复位沿检测实例 / Phase reset edge detector instance
    ePhase      : E_DL_PulsePhase;    // 相位状态机 / Phase state machine
    tHighTime   : TIME;               // 高电平持续 [ms] / High duration [ms]
    tLowTime    : TIME;               // 低电平持续 [ms] / Low duration [ms]
    tPeriodEff  : TIME;               // 钳位后周期 [ms] / Clamped period [ms]
    tPhasePt    : TIME;               // 当前相位定时器预设 [ms] / Preset of the current phase [ms]
    fDutyEff    : REAL;               // 钳位后占空比 [0..1] / Clamped duty [0..1]
    fPeriodMs   : REAL;               // 周期毫秒实数 [ms] / Period in milliseconds [ms]
    fHighMs     : REAL;               // 高相位毫秒实数 [ms] / High phase in milliseconds [ms]
    bParamBad   : BOOL;               // 参数钳位告警 / Parameter clamp warning
    bStateBad   : BOOL;               // 非法状态命中 / Illegal state hit
    bPhaseSwitched : BOOL;            // 本周期发生相位切换 / A phase switch happened this scan
    bRestartMask   : BOOL;            // 下一周期断开相位定时器一扫描（ET 归零）/ Drop the timer input for one scan
END_VAR
VAR CONSTANT
    DL_PULSE_PERIOD_MIN : TIME  := T#2MS;     // 周期下限 [ms]，至少两个任务周期可辨 / Min period [ms]
    DL_PULSE_PERIOD_MAX : TIME  := T#12H;     // 周期上限 [ms] / Max period [ms]
    DL_FLOAT_EPS        : REAL  := 1.0E-6;    // 浮点判零容差 / Float zero tolerance
END_VAR

(*------------------------------------------------------------------------------
 * 段 1｜无条件刷新区（红线 R7）：复位沿实例位于主体最前部，严禁进入 IF / CASE
 *      Unconditional refresh zone: the reset edge instance runs at the very top
 *-----------------------------------------------------------------------------*)
fbTrigReset(CLK := bPhaseReset);

(*------------------------------------------------------------------------------
 * 段 2｜占空比钳位（边界 B2）：越界钳位后继续运行并告警，与 0/1 的比较用容差
 *      Duty clamping: out-of-range values clamp and warn, comparisons use a tolerance
 *-----------------------------------------------------------------------------*)
bParamBad := FALSE;

IF fDutyCycle < 0.0 THEN
    fDutyEff  := 0.0;
    bParamBad := TRUE;
ELSIF fDutyCycle > 1.0 THEN
    fDutyEff  := 1.0;
    bParamBad := TRUE;
ELSE
    fDutyEff  := fDutyCycle;
END_IF

(*------------------------------------------------------------------------------
 * 段 3｜周期钳位（边界 B3）：下限防丢沿、上限防时间量溢出，两端都告警
 *      Period clamping: the lower bound prevents missed edges downstream
 *-----------------------------------------------------------------------------*)
IF tPeriod < DL_PULSE_PERIOD_MIN THEN
    tPeriodEff := DL_PULSE_PERIOD_MIN;
    bParamBad  := TRUE;
ELSIF tPeriod > DL_PULSE_PERIOD_MAX THEN
    tPeriodEff := DL_PULSE_PERIOD_MAX;
    bParamBad  := TRUE;
ELSE
    tPeriodEff := tPeriod;
END_IF

(*------------------------------------------------------------------------------
 * 段 4｜时长拆分（边界 B5/B9）：高相位时长由周期 × 占空比得出，低相位取差值
 *      Duration split: high = period x duty, low is the remainder
 *      先钳位高相位不超过整周期，杜绝换算误差造成的负重
 *      The high phase is clamped to the period so rounding can never go negative
 *-----------------------------------------------------------------------------*)
fPeriodMs := TIME_TO_REAL(tPeriodEff);
fHighMs   := fPeriodMs * fDutyEff;

IF fHighMs < 0.0 THEN
    fHighMs := 0.0;
ELSIF fHighMs > fPeriodMs THEN
    fHighMs := fPeriodMs;
END_IF

tHighTime := REAL_TO_TIME(fHighMs);
tLowTime  := tPeriodEff - tHighTime;

(*------------------------------------------------------------------------------
 * 段 5｜相位定时器刷新（边界 B1）：PT 由当前相位决定，IN 在复位与换相周期断开
 *      Phase timer refresh: PT follows the current phase, IN drops on reset and on a switch
 *      复位当周期 IN 为 FALSE 使 ET 立即清零，实现"从高相位起点重新起算"
 *      A FALSE IN on the reset scan clears ET so the high phase restarts from zero
 *      换相后必须再断一拍：标准定时器只在 IN 为 FALSE 时清 ET，
 *      仅改 PT 不会清零，ET 会带着上一相位的残值继续累加，
 *      低相位因此被缩短为一个扫描周期（v1.0.1 修复的正是此缺陷）
 *      A PT change never clears ET; without one off-scan the low phase collapses
 *-----------------------------------------------------------------------------*)
IF ePhase = eLow THEN
    tPhasePt := tLowTime;
ELSE
    tPhasePt := tHighTime;
END_IF

fbTonPhase(IN  := ((ePhase = eHigh) OR (ePhase = eLow)) AND bEnable
                  AND (NOT fbTrigReset.Q) AND (NOT bRestartMask),
           PT  := tPhasePt);

(*------------------------------------------------------------------------------
 * 段 6｜状态机（边界 B6/B7/B8）：禁用回首态，复位回高相位，相位期满互换
 *      State machine: disable parks at init, reset returns to high, expiry swaps
 *-----------------------------------------------------------------------------*)
bStateBad := FALSE;
bPhaseSwitched := FALSE;

IF NOT bEnable THEN
    (* 禁用：回首态并强制输出低；重新使能从高相位起步，不与外设中途相位错位 *)
    (* Disabled: park at init and force the output low; re-enable restarts at high *)
    ePhase := eInit;
ELSIF fbTrigReset.Q THEN
    (* 相位复位：本周期定时器已被清零，下一次调用从高相位重新计时 *)
    (* Phase reset: the timer is already cleared, the next call times the high phase *)
    ePhase := eHigh;
ELSE
    CASE ePhase OF

        eInit:
            (* 首态：使能后从高电平相位起步 *)
            (* Initial state: enter the high phase once enabled *)
            ePhase := eHigh;

        eHigh:
            (* 高相位期满：切换到低相位，并申请下一周期断拍使 ET 归零 *)
            (* High phase expired: switch to low and request one off-scan to clear ET *)
            IF fbTonPhase.Q THEN
                ePhase         := eLow;
                bPhaseSwitched := TRUE;
            END_IF

        eLow:
            (* 低相位期满：回到高相位，同样断拍一拍重新起算 *)
            (* Low phase expired: back to high with the same one-scan restart *)
            IF fbTonPhase.Q THEN
                ePhase         := eHigh;
                bPhaseSwitched := TRUE;
            END_IF

        eFault:
            (* 故障锁存：输出由段 7 强制低，等待禁用或复位 *)
            (* Fault latched: stage 7 forces the output low until disable or reset *)
            ePhase := eFault;

        ELSE
            (* 非法相位拦截：转故障并上报，不做隐式恢复 *)
            (* Illegal phase interception: go to fault and report, no implicit recovery *)
            ePhase    := eFault;
            bStateBad := TRUE;

    END_CASE;
END_IF

(*------------------------------------------------------------------------------
 * 段 7｜输出单一出口（边界 B4/B8）：恒低/恒高两态显式分支，不依赖相位机碰运气
 *      Single output outlet: degenerate duties take explicit branches
 *      占空比恰为 0 或 1 时若走相位机，会出现"进入高相位当周期即判期满"的毛刺
 *      Routing degenerate duties through the phase machine would create a one-scan glitch
 *-----------------------------------------------------------------------------*)
IF NOT bEnable THEN
    bPulseOut := FALSE;
ELSIF ABS(fDutyEff) <= DL_FLOAT_EPS THEN
    bPulseOut := FALSE;
ELSIF ABS(fDutyEff - 1.0) <= DL_FLOAT_EPS THEN
    bPulseOut := TRUE;
ELSIF ePhase = eHigh THEN
    bPulseOut := TRUE;
ELSE
    bPulseOut := FALSE;
END_IF

(*------------------------------------------------------------------------------
 * 段 8｜进度输出（边界 B9）：按相位累计 ET，除零前置判零 + 结果双向钳位
 *      Progress output: ET accumulated per phase, divide guard plus two-sided clamp
 *-----------------------------------------------------------------------------*)
IF fPeriodMs > DL_FLOAT_EPS THEN
    IF ePhase = eHigh THEN
        fProgress := TIME_TO_REAL(fbTonPhase.ET) / fPeriodMs;
    ELSIF ePhase = eLow THEN
        fProgress := (fHighMs + TIME_TO_REAL(fbTonPhase.ET)) / fPeriodMs;
    ELSE
        fProgress := 0.0;
    END_IF
ELSE
    fProgress := 0.0;
END_IF

IF fProgress < 0.0 THEN
    fProgress := 0.0;
ELSIF fProgress > 1.0 THEN
    fProgress := 1.0;
END_IF

(*------------------------------------------------------------------------------
 * 段 9｜故障码汇总：非法状态优先，其余为参数钳位告警
 *      Error aggregation: an illegal state outranks the parameter clamp warnings
 *-----------------------------------------------------------------------------*)
IF bStateBad THEN
    uErrorId := 16#0001_0005;
ELSIF bParamBad THEN
    uErrorId := 16#0001_0001;
ELSE
    uErrorId := 16#0000_0000;
END_IF

bError := (uErrorId <> 16#0000_0000);

(*------------------------------------------------------------------------------
 * 段 10｜换相断拍提交：本周期置的切换请求在下一周期生效并自动解除
 *      Switch mask commit: a switch raised this scan drops IN next scan and self-clears
 *      与顺控引擎的换步屏蔽同一范式：请求提交延后一拍，避免同周期自锁
 *      Same idiom as the sequencer's step mask: commit one scan later, never self-locking
 *-----------------------------------------------------------------------------*)
bRestartMask := bPhaseSwitched;
END_FUNCTION_BLOCK

(* ---- FB_DL_PulseSeqVerify.st ---- *)
(*==============================================================================
 * 组件名称 (Component)  : FB_DL_PulseSeqVerify
 * 所属子库 (Sublibrary) : DL_Base
 * 当前版本 (Version)    : 1.0.0
 * 兼容性 (Platform)     : CODESYS 3.5+ / TwinCAT 3 / 汇川 InoProShop / 施耐德 Machine Expert
 *                         仅依赖 Standard.library（TON / R_TRIG），零厂商私有库
 * 功能描述 (Function)   : 脉冲序列完整性校验。bStartCmd 上升沿武装并清零计数，
 *                         随后在开放窗口内对 bPulseIn 计数（实测 m），窗口关闭
 *                         条件 = 实测达到期望 n 或窗口超时 tWindow。收口时比对：
 *                         m = n → 序列完整 bSeqOk 单拍置位；m < n → 丢失判据
 *                         bSeqFail 置位并输出缺口数 nMissing = n - m；m > n
 *                         视为串扰/抖动超差同样判失败（缺失/多计双口径）。
 *                         步进电机丢步、流量脉冲丢失、编码器脉冲串完整性场景。
 * 来源标签 (Origin)     : 自研线（IEC 61131-3 标准语义的道莅防御性实现，clean-room）
 * 分工声明 (Pairing)    : PulseSeqVerify（序列完整性，本件）↔ EventCounter（无序
 *                         事件计数，既有件）：本件管「期望 n 与实测 m 的有序
 *                         比对与窗口收口」，不做无限累计计数；EventCounter 只
 *                         累计不比对、不判完整性。
 * 输出语义 (Fallback)   : 【R191】eIdle 相 → 全输出缺省零值；eFault 相 → 计数
 *                         与比对结果冻结保持末值，bError = TRUE；窗口运行中
 *                         失能 → 本轮作废、计数清零（作废语义在此声明）。
 * 组态闸 (Config gate)  : nPulseExpect < 1（无序列可验）或 tWindow <= T#0S
 *                         → 故障锁存（PT 为保持时长语义，非超时上限，R219 口径）。
 * 码位     (Codes)      : 按 R297 范式零 16# 码位硬编码；错误出口 BOOL+ENUM(eCause)，
 *                         码位待主控收口统一派号。
 * 红线自检 (Redline)    : 7 项红线已自检：R1 零全局 ✓｜R2 零物理地址 ✓｜R3 纯 IEC ✓
 *                         R4 组态闸/整型域防御（DINT 计数防回绕）✓
 *                         R5 双语同行注释 ✓｜R6 CASE 带 ELSE 兜底迁 eFault ✓
 *                         R7 TON/R_TRIG 段 0 无条件每拍刷新，各实例单用途 ✓
 * 验收向量 (Acceptance) : V1 期望 100 实测恰 100 → bSeqOk 单拍 TRUE；
 *                         V2 期望 100 实测 97 → bSeqFail=TRUE，nMissing=3；
 *                         V3 期望 100 窗口到时仅 40 → bSeqFail，nMissing=60；
 *                         V4 复位沿清全部计数与锁存 → 上电回夹防线（R268）。
 * 修订历史 (Revision)   : 2026-11-20  v1.0.0  R49 首版（批 1 · 序号 4）
 *==============================================================================*)
TYPE E_DL_PsvState :
(
    eIdle   := 0,                            (* 待武装（输出缺省） / Idle, disarmed *)
    eArmed  := 10,                           (* 计数窗口开放中 / Counting window open *)
    eDone   := 20,                           (* 本轮收口完成，结果保持 / Round closed, result held *)
    eFault  := 90                            (* 故障锁存相 / Fault latched phase *)
);
END_TYPE

TYPE E_DL_PsvCause :
(
    eNone       := 0,                        (* 无故障成因 / No cause *)
    eCfgIllegal := 1,                        (* 组态非法：期望数/窗口越域 / Illegal config *)
    ePhaseBad   := 2                         (* 非法相位兜底 / Illegal phase fallback *)
);
END_TYPE

FUNCTION_BLOCK FB_DL_PulseSeqVerify
VAR_INPUT
    bPulseIn    : BOOL := FALSE;             (* 被校验脉冲输入（内部取上升沿）[-] / Pulse input to verify *)
    nPulseExpect: DINT := 100;               (* 期望脉冲数 n，域 >= 1 [个] / Expected pulse count, domain >= 1 *)
    tWindow     : TIME := T#10S;             (* 计数开放窗口保持时长（收口时限语义）[ms] / Counting window hold time *)
    bStartCmd   : BOOL := FALSE;             (* 启动命令，上升沿武装本轮并清零计数 [-] / Start command, rising edge arms round *)
    bEnable     : BOOL := TRUE;              (* 校验使能，运行中失能则本轮作废清零 [-] / Enable, disable aborts current round *)
    bReset      : BOOL := FALSE;             (* 复位命令，上升沿清全部内部状态 [-] / Reset, rising edge clears all internal state *)
END_VAR
VAR_OUTPUT
    nPulseMeas  : DINT;                      (* 本轮实测脉冲数 m（收口后保持）[个] / Measured pulse count this round *)
    nMissing    : DINT;                      (* 缺口数 = n - m（多计为负值），收口后保持 [个] / Missing count, negative on overrun *)
    bSeqOk      : BOOL;                      (* 本轮序列完整单拍位（m = n 收口拍置位）[-] / Round-complete single-scan flag *)
    bSeqFail    : BOOL;                      (* 本轮序列不完整锁存位（收口至复位沿）[-] / Round-incomplete latch until reset *)
    bCounting   : BOOL;                      (* 窗口开放中指示 [-] / Window-open indicator *)
    eState      : E_DL_PsvState;             (* 状态出口 / State outlet *)
    eCause      : E_DL_PsvCause;             (* 故障成因出口（R190 归因唯一） / Fault cause outlet *)
    bError      : BOOL;                       (* 故障锁存标志 [-] / Fault latch flag *)
END_VAR
VAR
    _eState   : E_DL_PsvState := E_DL_PsvState.eIdle;      (* 内部相位（CASE 唯一写入目标） / Internal phase *)
    _eCause   : E_DL_PsvCause := E_DL_PsvCause.eNone;      (* 故障成因锁存量 / Latched cause *)
    rtPulse   : R_TRIG;                     (* 脉冲上升沿实例，段 0 无条件调用 / Pulse rising edge *)
    rtStart   : R_TRIG;                     (* 启动上升沿实例，段 0 无条件调用 / Start rising edge *)
    rtReset   : R_TRIG;                     (* 复位上升沿实例，段 0 无条件调用 / Reset rising edge *)
    tonWindow : TON;                        (* 窗口计时，IN 由相位派生，段 0 无条件调用 / Window timer *)
    _nCount   : DINT;                       (* 实测计数锁存（本轮累计量）[个] / Measured count latch *)
    _bFault   : BOOL;                       (* 故障锁存位 / Latched fault bit *)
    _bCfgBad  : BOOL;                       (* 组态非法当拍量 / Illegal config this scan *)
    _bResult  : BOOL;                       (* 本轮收口判据：TRUE 完整 / FALSE 不完整 / Round verdict latch *)
END_VAR

(* —— 段 0：当拍判据派生 + 实例无条件周期刷新（R228A） —— *)
_bCfgBad := (nPulseExpect < 1) OR (tWindow <= T#0S);       (* 组态闸：期望数与窗口越域 / Config gate *)
rtPulse(CLK := bPulseIn);                                   (* 脉冲沿每拍必调 / Pulse edge every scan *)
rtStart(CLK := bStartCmd);                                  (* 启动沿每拍必调 / Start edge every scan *)
rtReset(CLK := bReset);                                     (* 复位沿每拍必调 / Reset edge every scan *)
tonWindow(IN := _eState = E_DL_PsvState.eArmed, PT := tWindow);   (* 窗口计时随相位派生 / Window timer phase-derived *)

(* —— 段 1：单拍量预清零（锁存量与实例不入清单，R107） —— *)
bSeqOk := FALSE;                                            (* 完整单拍位预清，唯一分支置位 / Complete pulse preset *)

(* —— 段 2：复位沿处理（作用域：清锁存 + 清计数 + 清结果 + 迁 eIdle，R283 逐项声明） —— *)
IF rtReset.Q THEN
    _bFault := FALSE;                                       (* 清故障锁存 / Clear fault latch *)
    _eCause := E_DL_PsvCause.eNone;                         (* 清成因 / Clear cause *)
    _nCount := 0;                                           (* 清实测计数 / Clear count *)
    _bResult := FALSE;                                      (* 清结果锁存 / Clear verdict latch *)
    nPulseMeas := 0;                                        (* 清输出计数镜像 / Clear output count *)
    nMissing := 0;                                          (* 清缺口输出 / Clear missing output *)
    bSeqFail := FALSE;                                      (* 清失败锁存 / Clear fail latch *)
    _eState := E_DL_PsvState.eIdle;                         (* 迁待武装相 / Back to idle *)
END_IF

(* —— 段 3：组态闸故障锁存（赋值 3 行内置 bError，R45 配对；锁存至复位沿，R189） —— *)
IF _bCfgBad AND NOT _bFault THEN
    _bFault := TRUE;                                        (* 锁存故障位 / Latch fault *)
    _eCause := E_DL_PsvCause.eCfgIllegal;                   (* 成因：组态非法 / Cause: illegal config *)
    _eState := E_DL_PsvState.eFault;                        (* 同步迁故障相 / Migrate to fault *)
END_IF

(* —— 段 4：CASE 主状态机（ELSE 兜底迁 eFault，红线 6） —— *)
CASE _eState OF
    E_DL_PsvState.eIdle:                                    (* 待武装相 / Idle *)
        IF rtStart.Q AND bEnable AND NOT _bFault THEN
            _nCount := 0;                                   (* 武装清零本轮计数 / Arm clears count *)
            _eState := E_DL_PsvState.eArmed;                (* 进入计数窗口 / Enter armed *)
        END_IF
    E_DL_PsvState.eArmed:                                   (* 计数窗口相 / Armed *)
        IF NOT bEnable THEN                                 (* 运行中失能：本轮作废清零（声明语义） / Disable aborts round *)
            _nCount := 0;                                   (* 作废清计数 / Abort clears count *)
            _eState := E_DL_PsvState.eIdle;                 (* 回待武装 / Back to idle *)
        ELSIF rtPulse.Q THEN
            _nCount := _nCount + 1;                         (* 脉冲计数（DINT 域，窗口时限天然防回绕） / Increment count *)
        END_IF
        IF _eState = E_DL_PsvState.eArmed AND (_nCount >= nPulseExpect OR tonWindow.Q) THEN
            nPulseMeas := _nCount;                          (* 收口：实测镜像 / Close round: mirror count *)
            nMissing := nPulseExpect - _nCount;             (* 缺口数（多计为负） / Missing, negative on overrun *)
            _bResult := (_nCount = nPulseExpect);           (* 完整判据：恰等（整型用等值比较合法） / Verdict: exact equality *)
            bSeqOk := _bResult;                             (* 完整单拍位 / Complete pulse *)
            bSeqFail := NOT _bResult;                       (* 失败锁存至复位沿 / Fail latch until reset *)
            _eState := E_DL_PsvState.eDone;                 (* 迁收口相 / Enter done *)
        END_IF
    E_DL_PsvState.eDone:                                    (* 收口保持相：结果冻结，等下一轮武装或复位 / Done: hold result *)
        IF rtStart.Q AND bEnable AND NOT _bFault THEN       (* 新一轮武装重启 / New round re-arms *)
            _nCount := 0;                                   (* 清本轮计数 / Clear count *)
            bSeqFail := FALSE;                              (* 清上一轮失败锁存 / Clear previous fail latch *)
            _eState := E_DL_PsvState.eArmed;                (* 进入计数窗口 / Enter armed *)
        END_IF
    E_DL_PsvState.eFault:                                   (* 故障相：冻结保持，仅复位沿出 / Fault: frozen *)
        ;                                                   (* 锁存回放（R28） / Replay from latch *)
    ELSE                                                    (* 非法相位兜底迁安全态 / Illegal phase fallback *)
        _eState := E_DL_PsvState.eFault;                    (* 迁故障相 / To fault *)
        _bFault := TRUE;                                    (* 同步锁存 / Latch *)
        _eCause := E_DL_PsvCause.ePhaseBad;                 (* 成因：非法相位 / Cause: illegal phase *)
END_CASE

(* —— 段 5：出口映射（bError/eState 同源，R191） —— *)
bCounting := (_eState = E_DL_PsvState.eArmed);              (* 窗口开放指示 / Window-open indicator *)
nPulseMeas := _nCount;                                      (* 实测计数实时镜像（窗口中也可见） / Live count mirror *)
bError := _bFault;                                          (* 故障标志镜像 / Fault flag mirror *)
eState := _eState;                                          (* 状态出口 / State outlet *)
eCause := _eCause;                                          (* 成因出口 / Cause outlet *)
END_FUNCTION_BLOCK

(* ---- FB_DL_PulseStretch.st ---- *)
(*
    FB_DL_PulseStretch —— 脉冲展宽（最小脉宽保持）
    ------------------------------------------------------------------
    分类      : DL_Base / Signal
    前缀      : FB_DL_
    版本      : 1.0.0
    溯源      : T0-2 定时器族变体（ADR：TON 语义 + 最小脉宽工况）；
                T1-1 OSCAT Basic 信号整形惯例为次源，只借「最小脉宽保持」这一
                整形分类事实，不复制任何函数体；clean-room 重写，未复制任何
                闭源厂商源码，参考实现仅限 MIT/Apache 许可
    平台      : 纯 IEC 61131-3，CODESYS V3.5+ / TwinCAT 3 / InoProShop 通用
    作者      : 道莅代码库 · PLC编程专家（R18）
    ------------------------------------------------------------------
    功能说明  : 现场窄脉冲（< 执行机构最小响应时间）会被下游设备吃掉，本件把输出
                保持到满足最小脉宽 tMinPulse 才释放；双模：可重触发（保持期内新沿
                重新计时）与不可重触发（计时不重启）；
                tMinPulse 非法（0 或 < 1 ms）退化为直通，绝不把 TON 置于非法 PT；
                tMinPulse 超上限先钳位到 10 s 再进定时器；
                与 FB_DL_SignalDebounce（去抖）职责互补，本件不做滤波。
    错误码    : 16#0001_0237 tMinPulse 超上限已钳位到 10 s——信息级，正常防御
                16#0001_0238 预留禁用（信息级，不得挪用）
                16#0001_0309 tMinPulse 非法（< 1 ms 或 0）——故障级，本拍退化为直通
                16#0001_030A 预留禁用（故障级，不得挪用）
                16#0001_030B 预留禁用（故障级，不得挪用）
    码位总账  : 16#0001_0237 用 / 16#0001_0238 预留 ｜ 16#0001_0309 用 / 16#0001_030A 预留 / 16#0001_030B 预留
    状态机    : 无 CASE，保持期由 TON 的 ET 与单比特 bHoldActive 承载，非法状态不可能出现
    采样约定  : fbTrigIn / fbHold 两个实例在本体首部无条件调用，ET 不会冻结；
                输入脉冲短于一个扫描周期不可见（与库内 SineGenerator 同口径），
                低于任务频率一半的脉冲必须先经硬件或高速任务采样。
    修订记录  : 2026-11-16 v1.0.0 首次入库（R18）
*)
FUNCTION_BLOCK FB_DL_PulseStretch
VAR_INPUT
    bEnable        : BOOL;                     // 使能，FALSE 输出立即复位 / enable, FALSE resets the output immediately
    bIn            : BOOL;                     // 脉冲输入，已在别处去抖时可直接连接 / pulse input, connect directly when debounced upstream
    tMinPulse      : TIME := T#50MS;           // 最小输出脉宽 [ms]，范围 1~10000，0 非法 / minimum output pulse width [ms], range 1~10000, 0 illegal
    bRetriggerable : BOOL := TRUE;             // TRUE 重触发 / FALSE 保持期内不重启计时 / TRUE retriggerable, FALSE keeps the running timer
END_VAR
VAR_OUTPUT
    bOut        : BOOL;                        // 展宽后的输出 / stretched output
    bStretching : BOOL;                        // 正在展宽（保持期） / currently stretching (hold phase)
    tRemain     : TIME;                        // 保持期剩余时间 [ms] / remaining hold time [ms]
    uStretchCnt : UDINT;                       // 累计展宽次数，饱和计数 [次] / accumulated stretch count, saturating [times]
    eErr        : UDINT;                       // 错误码，0=正常 / error id, 0=ok
    bError      : BOOL;                        // 故障标志，eErr 为故障级时 TRUE / error flag, TRUE on fault-level eErr
END_VAR
VAR
    fbTrigIn    : R_TRIG;                      // 输入上升沿检测实例，本体首部无条件刷新 / input rising edge instance, refreshed unconditionally
    fbHold      : TON;                         // 保持期定时器实例，本体首部无条件刷新 / hold phase timer, refreshed unconditionally
    bHoldActive : BOOL;                        // 保持期有效位，下一拍作为定时器 IN / hold phase active bit, fed to the timer input next cycle
    bPassThru   : BOOL;                        // 直通退化标志，脉宽参数非法时为 TRUE / pass-through fallback flag, TRUE when the width parameter is illegal
    bRestart    : BOOL;                        // 重触发请求标志，单拍 / retrigger request flag, single cycle
    bInit       : BOOL := FALSE;               // 首扫标志，初值 FALSE，判据 NOT bInit / first-scan flag, initial FALSE, tested with NOT
    tEffMin     : TIME := T#50MS;              // 生效最小脉宽，钳位后进入定时器 [ms] / effective minimum width fed to the timer [ms]
    tRem        : TIME;                        // 剩余时间中间量 [ms] / remaining time intermediate [ms]
END_VAR
VAR CONSTANT
    DL_STRETCH_MIN     : TIME := T#1MS;        // 最小脉宽下限 [ms] / lower bound of the pulse width [ms]
    DL_STRETCH_MAX     : TIME := T#10S;        // 最小脉宽上限 [ms] / upper bound of the pulse width [ms]
    DL_STRETCH_CNT_MAX : UDINT := 16#FFFF_FFFE;// 展宽计数饱和值，防回绕 [次] / stretch counter saturation value, no wrap-around [times]
END_VAR

// 段 1｜输出与错误状态预置 / segment 1, preset outputs and error status
eErr := 0;                                     // 预置无错误 / preset no error
bError := FALSE;                               // 预置无故障 / preset no fault
tRemain := T#0MS;                              // 剩余时间先归零 / remaining time to zero
bPassThru := FALSE;                            // 直通标志先清 / clear the pass-through flag

// 段 2｜首扫初始化（初值 FALSE，判据 NOT bInit）/ segment 2, first-scan initialisation
IF NOT bInit THEN
    bHoldActive := FALSE;                      // 首扫不得处于保持期 / no hold phase may survive the first scan
    uStretchCnt := 0;                          // 计数从 0 起 / counter starts at zero
    bInit := TRUE;                             // 首扫只做一次 / first scan runs once only
END_IF

// 段 3｜脉宽参数闸：先判非法（退化直通），再判超限（钳位后进定时器）/ segment 3, pulse width parameter gate
tEffMin := tMinPulse;                          // 默认沿用输入值 / default to the input value
IF tMinPulse < DL_STRETCH_MIN THEN
    tEffMin := DL_STRETCH_MIN;                 // 定时器必须拿到合法 PT / the timer must receive a legal preset
    bPassThru := TRUE;                         // 退化为直通 / degrade to pass-through
    eErr := 16#0001_0309;                      // 脉宽非法故障码 / illegal pulse width fault id
    bError := TRUE;                            // 置故障标志 / raise the error flag
ELSIF tMinPulse > DL_STRETCH_MAX THEN
    tEffMin := DL_STRETCH_MAX;                 // 超上限先钳位 / clamp to the upper bound first
    eErr := 16#0001_0237;                      // 钳位提示（信息级不置故障）/ clamp hint, info level never raises a fault
END_IF

// 段 4｜边沿与定时器实例无条件周期刷新（红线：ET 绝不冻结）/ segment 4, unconditional refresh of the edge and timer instances
fbTrigIn(CLK := bIn);                          // 输入沿 / input edge
fbHold(IN := bHoldActive, PT := tEffMin);      // 保持期定时器，本拍 IN 取上一拍有效位 / hold timer, input uses the previous cycle value

// 段 5｜失能闸：立即复位输出并清保持期 / segment 5, enable gate resets the output immediately
IF NOT bEnable THEN
    bHoldActive := FALSE;                      // 清保持期 / clear the hold phase
    bOut := FALSE;                             // 输出复位 / reset the output
    bStretching := FALSE;                      // 非展宽态 / not stretching
    tRemain := T#0MS;                          // 剩余时间归零 / remaining time to zero
    RETURN;                                    // 失能即出口 / disabled is the exit
END_IF

// 段 6｜直通退化：参数非法时不进定时器 / segment 6, pass-through fallback bypasses the timer
IF bPassThru THEN
    bHoldActive := FALSE;                      // 直通不维持保持期 / no hold phase in pass-through mode
    bOut := bIn;                               // 输出等于输入 / output equals input
    bStretching := FALSE;                      // 非展宽态 / not stretching
    tRemain := T#0MS;                          // 剩余时间归零 / remaining time to zero
    RETURN;                                    // 直通即出口 / pass-through is the exit
END_IF

// 段 7｜重触发判定：本拍先掉 IN 一拍以让 TON 复位，下一拍重新计时 / segment 7, retrigger drops the timer input for one cycle
bRestart := fbTrigIn.Q AND bRetriggerable AND bHoldActive; // 仅可重触发且已在保持期时成立 / only in retriggerable mode while already holding
IF bIn THEN
    bHoldActive := TRUE;                       // 输入到来即进入保持期 / an active input starts the hold phase
END_IF
IF bRestart THEN
    bHoldActive := FALSE;                      // 单拍掉 IN，ET 归零，下一拍重新计时 / drop the input for one cycle so ET restarts next cycle
END_IF

// 段 8｜保持期满释放 / segment 8, release after the hold phase expires
IF fbHold.Q THEN
    bHoldActive := FALSE;                      // 期满释放 / release when the preset is reached
END_IF

// 段 9｜展宽次数统计（饱和，不回绕）/ segment 9, stretch counter with saturation
IF fbTrigIn.Q AND (NOT bRestart) THEN
    IF uStretchCnt < DL_STRETCH_CNT_MAX THEN
        uStretchCnt := uStretchCnt + 1;        // 饱和加一，绝不回绕 / saturating increment, never wraps
    END_IF
END_IF

// 段 10｜输出与剩余时间：剩余时间用 PT 减 ET，ET 不小于 PT 时归零 / segment 10, output and remaining time
bStretching := bHoldActive;                    // 保持期镜像 / hold phase mirror
bOut := bIn OR bHoldActive;                    // 输入为真或仍在保持期则输出为真 / TRUE while the input is on or the hold phase runs
IF fbHold.ET < tEffMin THEN
    tRem := tEffMin - fbHold.ET;               // 剩余 = 最小脉宽减已保持 / remaining = preset minus elapsed
ELSE
    tRem := T#0MS;                             // 已到期，剩余归零 / expired, remaining is zero
END_IF
tRemain := tRem;                               // 对外镜像 / publish the remaining time
END_FUNCTION_BLOCK

(* ---- FB_DL_PulseTrainDecoder.st ---- *)
(*
  Name        : FB_DL_PulseTrainDecoder
  Category    : DL_Base
  Version     : 1.0.0
  Purpose     : 脉冲串解码：统计脉冲总数，按脉宽宽/窄逐位移入编码字，间隔超窗即判整字完成并锁存输出（编码旋钮/拨码开关读入）；/ Pulse-train decoder: counts pulses, shifts wide/narrow pulse bits into a code word, and latches the word when the inter-pulse gap window elapses (encoder knob / DIP-switch read-in)
  溯源        : 借 t2-1-lgf-bit-logic 的分类/参数域组织，clean-room 实现
  Boundary    : ① 组态闸：宽脉冲阈/间隔窗任一 <= 0 或间隔窗 <= 宽阈 → 锁存故障（间隔窗必须显著大于宽阈才可区分字间隔与位间隔）；
                ② 位容量 16 位：位满后继续收到的脉冲只计数不再移位（防溢出回绕破坏编码）；
                ③ 宽窄判据用「脉宽 TON（IN := bPulse）在下降沿读上拍 Q」的上一拍口径，段 0 无 IF 包裹刷新；
                ④ 间隔判定 TON 串 eRx 相位闸（族③），字完成沿由 R_TRIG 提取（R187 两段式）；
                ⑤ nCode/nBits 在 eDone 相保持（锁存副本），直到下一个字首脉冲或复位才刷新（族② 保持语义）；
                ⑥ 本件只解码，不执行旋钮联动逻辑（属主边界）。
*)
TYPE E_DL_PtdState :
(
    eIdle := 0,                              (* 未使能 / Disabled *)
    eRx   := 10,                             (* 收码中（位流移入） / Receiving *)
    eDone := 20,                             (* 字完成（保持编码） / Word complete, held *)
    eFault:= 90                              (* 故障锁存相 / Fault latched *)
);
END_TYPE

TYPE E_DL_PtdCause :
(
    eNone       := 0,                        (* 无故障成因 / No cause *)
    eCfgIllegal := 1,                        (* 组态非法：宽阈/间隔窗越域 / Illegal config *)
    ePhaseBad   := 2                         (* 非法相位兜底 / Illegal phase fallback *)
);
END_TYPE

FUNCTION_BLOCK FB_DL_PulseTrainDecoder
VAR_INPUT
    bPulse   : BOOL := FALSE;                (* 脉冲串输入电平 [-] / Pulse-train input *)
    tWideMin : TIME := T#30MS;               (* 宽脉冲下限（脉宽 >= 此值判 1），域 > T#0S [ms] / Wide-pulse threshold, > 0 *)
    tGapMax  : TIME := T#300MS;              (* 位间隔窗（间隔超此值判整字结束），域 > 宽阈 [ms] / Bit-gap window, > wide threshold *)
    bEnable  : BOOL := TRUE;                 (* 解码使能 [-] / Enable *)
    bReset   : BOOL := FALSE;                (* 复位命令，上升沿清计数与编码 [-] / Reset command *)
END_VAR
VAR_OUTPUT
    nPulseCnt: UDINT;                        (* 累计脉冲总数（饱和）[个] / Total pulse count, saturated *)
    nCode    : UDINT;                        (* 最近完成字的编码值（eDone 相保持）[-] / Last completed word code, held *)
    nBits    : INT;                          (* 最近完成字位数（eDone 相保持）[位] / Last completed word bit count, held *)
    bWordDone: BOOL;                         (* 字完成单拍脉冲 [-] / Word-complete single-scan pulse *)
    bRxOn    : BOOL;                         (* 收码进行中电平（eRx 相为 TRUE）[-] / Receiving level *)
    eState   : E_DL_PtdState;                (* 状态出口 / State outlet *)
    eCause   : E_DL_PtdCause;                (* 故障成因出口（R190 归因唯一） / Fault cause outlet *)
    bError   : BOOL;                         (* 故障锁存标志 [-] / Fault latch flag *)
END_VAR
VAR
    _eState  : E_DL_PtdState := E_DL_PtdState.eIdle;     (* 内部相位（CASE 唯一写入目标） / Internal phase *)
    _eCause  : E_DL_PtdCause := E_DL_PtdCause.eNone;     (* 故障成因锁存量 / Latched cause *)
    rtPulse  : R_TRIG;                       (* 脉冲上升沿实例，段 0 无条件调用 / Pulse rising edge *)
    rtFall   : R_TRIG;                       (* 脉冲下降沿实例，段 0 无条件调用 / Pulse falling edge *)
    rtGap    : R_TRIG;                       (* 间隔窗到点沿实例，段 0 无条件调用 / Gap-elapsed edge *)
    rtReset  : R_TRIG;                       (* 复位沿实例，段 0 无条件调用 / Reset edge instance *)
    tonWidth : TON;                          (* 脉宽测量计时器（IN := bPulse，下降沿读上拍 Q） / Pulse-width timer *)
    tonGap   : TON;                          (* 位间隔窗计时器（IN 串 eRx 相位） / Bit-gap timer *)
    _bFault  : BOOL;                         (* 故障锁存位 / Latched fault bit *)
    _bCfgBad : BOOL;                         (* 组态非法当拍量 / Illegal config this scan *)
    _bWide   : BOOL;                         (* 当前位宽窄当拍量（宽 = TRUE）[-] / Current bit wide flag *)
    _nCodeI  : UDINT;                        (* 收码移位寄存器内部量 [-] / Code shift register internal *)
    _nBitsI  : INT;                          (* 收码位数内部量 [位] / Bit count internal *)
    _bDoneC  : BOOL;                         (* 字完成内部单拍量（出口统一映射，R187） / Word-done internal pulse *)
END_VAR
VAR CONSTANT
    DL_PTD_CNTMAX : UDINT := 4294967295;     (* 脉冲计数饱和上限（R28）[-] / Pulse count saturation cap *)
    DL_PTD_BITMAX : INT   := 16;             (* 编码位容量上限（UDINT 移位安全域）[位] / Bit capacity limit *)
END_VAR

(* —— 段 0：当拍判据派生 + 实例无条件刷新（R228A；R_TRIG/TON 全在段 0，无 IF 包裹） —— *)
_bCfgBad := NOT (tWideMin > T#0S)                                              (* 宽脉冲阈正域闸 / Wide threshold gate *)
            OR NOT (tGapMax > T#0S)                                            (* 间隔窗正域闸 / Gap window gate *)
            OR (tGapMax <= tWideMin);                                          (* 间隔窗须大于宽阈（防位间隔误判字结束） / Gap window above wide threshold *)
rtPulse(CLK := bPulse);                                                        (* 上升沿每拍必调 / Rising edge every scan *)
rtFall(CLK := NOT bPulse);                                                     (* 下降沿每拍必调 / Falling edge every scan *)
rtReset(CLK := bReset);                                                        (* 复位沿每拍必调 / Reset edge every scan *)
tonWidth(IN := bPulse, PT := tWideMin);                                        (* 脉宽测量（下降沿读上拍 Q = 本脉冲是否够宽，边界③） / Width timer, prior-scan read at fall *)
tonGap(IN := (_eState = E_DL_PtdState.eRx) AND NOT bPulse, PT := tGapMax);     (* 位间隔窗（串 eRx 相位闸，族③） / Gap timer with phase gate *)
rtGap(CLK := tonGap.Q);                                                        (* 间隔窗到点沿每拍必调 / Gap edge every scan *)
_bWide := tonWidth.Q;                                                          (* 当前脉宽是否达宽阈（上一拍口径） / Current bit wide verdict *)

(* —— 段 1：单拍量预清零（R107） —— *)
_bDoneC := FALSE;                                                              (* 字完成内部量预清 / Word-done preset *)
bWordDone := FALSE;                                                            (* 字完成出口预清 / Word-done outlet preset *)
bRxOn := FALSE;                                                                (* 收码电平预清 / Rx level preset *)

(* —— 段 2：复位沿处理（作用域：清故障 + 清计数 + 清编码 + 迁 eIdle，R283 逐项声明） —— *)
IF rtReset.Q THEN
    _bFault := FALSE;                                                          (* 清故障锁存 / Clear fault *)
    _eCause := E_DL_PtdCause.eNone;                                            (* 清成因 / Clear cause *)
    nPulseCnt := 0;                                                            (* 清脉冲总数 / Clear pulse count *)
    nCode := 0;                                                                (* 清编码出口 / Clear code outlet *)
    nBits := 0;                                                                (* 清位数出口 / Clear bits outlet *)
    _nCodeI := 0;                                                              (* 清移位寄存器 / Clear shift register *)
    _nBitsI := 0;                                                              (* 清位数内部量 / Clear bit count internal *)
    _eState := E_DL_PtdState.eIdle;                                            (* 迁未使能相 / Back to idle *)
END_IF

(* —— 段 3：组态故障锁存（锁存至复位沿，R189） —— *)
IF _bCfgBad AND NOT _bFault THEN
    _bFault := TRUE;                                                           (* 锁存故障位 / Latch fault *)
    _eCause := E_DL_PtdCause.eCfgIllegal;                                      (* 成因：组态非法 / Cause: illegal config *)
    _eState := E_DL_PtdState.eFault;                                           (* 同步迁故障相 / Migrate to fault *)
END_IF

(* —— 段 4：CASE 主状态机（ELSE 兜底迁 eFault，红线 6） —— *)
CASE _eState OF
    E_DL_PtdState.eIdle:                                                       (* 未使能：不解码，出口确定值 / Disabled *)
        nPulseCnt := 0;                                                        (* 失能清脉冲总数 / Clear pulse count *)
        nCode := 0;                                                            (* 失能清编码出口 / Clear code outlet *)
        nBits := 0;                                                            (* 失能清位数出口 / Clear bits outlet *)
        _nCodeI := 0;                                                          (* 失能清移位寄存器 / Clear shift register *)
        _nBitsI := 0;                                                          (* 失能清位数内部量 / Clear bit count internal *)
        IF bEnable AND NOT _bFault THEN
            _eState := E_DL_PtdState.eRx;                                      (* 使能进入收码 / Enter receiving *)
        END_IF
    E_DL_PtdState.eRx:                                                         (* 收码相：位流移入 + 间隔判字 / Receiving *)
        IF NOT bEnable THEN
            _eState := E_DL_PtdState.eIdle;                                    (* 失能回未使能 / Back to idle *)
        ELSE
            IF rtPulse.Q THEN                                                  (* 字首脉冲：清移位寄存器重收新字 / First pulse of a word: clear register *)
                _nCodeI := 0;                                                  (* 移位寄存器清零 / Register clear *)
                _nBitsI := 0;                                                  (* 位数清零 / Bit count clear *)
            END_IF
            IF rtPulse.Q THEN                                                  (* 脉冲总数计数（与移位独立） / Total pulse count *)
                IF nPulseCnt < DL_PTD_CNTMAX THEN
                    nPulseCnt := nPulseCnt + 1;                                (* 净额 +1（饱和防回绕，R28） / Net +1, saturated *)
                END_IF
            END_IF
            IF rtFall.Q THEN                                                  (* 脉冲下降沿：本位宽窄已定，移入寄存器 / Bit settle at fall: shift in *)
                IF _nBitsI < DL_PTD_BITMAX THEN
                    _nCodeI := _nCodeI * 2;                                    (* 左移一位（位容量内，无溢出） / Shift left one bit *)
                    IF _bWide THEN
                        _nCodeI := _nCodeI + 1;                                (* 宽脉冲：该位为 1 / Wide bit: 1 *)
                    END_IF
                    _nBitsI := _nBitsI + 1;                                    (* 位数递进 / Bit count advance *)
                END_IF                                                         (* 位满后只计数不移位（边界②） / Beyond capacity: count only *)
            END_IF
            IF rtGap.Q THEN                                                    (* 间隔窗到点：整字结束 / Gap elapsed: word end *)
                IF _nBitsI > 0 THEN                                            (* 至少收到位才算有效字 / Word valid only with bits *)
                    nCode := _nCodeI;                                          (* 编码出口（锁存副本，eDone 相保持） / Code outlet, held *)
                    nBits := _nBitsI;                                          (* 位数出口（锁存副本） / Bits outlet, held *)
                    _bDoneC := TRUE;                                           (* 字完成内部置位（出口统一映射，R187） / Word-done internal *)
                END_IF
                _nCodeI := 0;                                                  (* 寄存器清零（下字重收） / Register clear *)
                _nBitsI := 0;                                                  (* 位数清零 / Bit count clear *)
                IF _bDoneC THEN
                    _eState := E_DL_PtdState.eDone;                            (* 有效字完成迁保持相 / To done on valid word *)
                END_IF
            END_IF
        END_IF
    E_DL_PtdState.eDone:                                                       (* 保持相：编码保持至下字首脉冲 / Done: hold code *)
        IF NOT bEnable THEN
            _eState := E_DL_PtdState.eIdle;                                    (* 失能回未使能 / Back to idle *)
        ELSIF rtPulse.Q THEN                                                   (* 下一个字首脉冲：回收码相重收 / Next word first pulse: back to rx *)
            _nCodeI := 0;                                                      (* 移位寄存器清零 / Register clear *)
            _nBitsI := 0;                                                      (* 位数清零 / Bit count clear *)
            _eState := E_DL_PtdState.eRx;                                      (* 回收码相 / Back to receiving *)
        END_IF
    E_DL_PtdState.eFault:                                                      (* 故障相：冻结保持末值，仅复位沿出 / Fault *)
        ;                                                                      (* 锁存回放（R28） / Replay from latch *)
    ELSE                                                                       (* 非法相位兜底迁安全态 / Illegal phase fallback *)
        _eState := E_DL_PtdState.eFault;                                       (* 迁故障相 / To fault *)
        _bFault := TRUE;                                                       (* 同步锁存 / Latch *)
        _eCause := E_DL_PtdCause.ePhaseBad;                                    (* 成因：非法相位 / Cause: illegal phase *)
END_CASE

(* —— 段 5：出口映射（内部 _b* → 输出，R187；名实双出口，R191） —— *)
bWordDone := _bDoneC;                                                          (* 字完成单拍出口 / Word-done single-scan outlet *)
bRxOn := (_eState = E_DL_PtdState.eRx);                                        (* 收码电平出口（相位镜像，R191） / Rx level outlet *)
bError := _bFault;                                                             (* 故障标志镜像 / Fault flag mirror *)
eState := _eState;                                                             (* 状态出口 / State outlet *)
eCause := _eCause;                                                             (* 成因出口 / Cause outlet *)
END_FUNCTION_BLOCK

(* ---- FB_DL_PulseWidthFilter.st ---- *)
(*
    组件名称 : FB_DL_PulseWidthFilter
    所属子库 : DL_Base
    当前版本 : 1.0.1
    兼 容 性 : CODESYS V3.5+ / TwinCAT 3 / 汇川 InoProShop；仅依赖 Standard.library
    功能描述 : 窄脉冲抑制，脉宽小于 tMinWidth 的整段脉冲不出现在输出上，合格脉冲的宽度不失真。
              取舍 ①（本件最容易写错的地方）：必须是「双侧确认窗」—— 上升沿与下降沿各用一只 TON 确认，
              输出相对输入整体滞后 tMinWidth。若只延迟上升沿（单侧确认），每个合格脉冲都会被削掉
              tMinWidth 的宽度，长信号看着正常、短脉冲悄悄变形，是现场最难查的一类错。
              本件用 fbOnDelay 确认高电平、fbOffDelay 确认低电平，两只看守各自一侧，于是宽度守恒。
              取舍 ②：窄脉冲「整段吞掉」而不是「压窄」—— 输出只在输入稳定维持 tMinWidth 后才跟随，
              未维持到确认完成的电平从来不落到输出上，抑制计数在「输入已回落但确认未完成」那拍递增。
              取舍 ③：失能即直通（bOut := bIn）—— 旁路时不得留门控残影；两只看守定时器的 IN 都串入 bEnable，
              保证失能期间它们同步复位，重新使能时从零开始确认，不会带着旧完成位直接放行。
              取舍 ④：与 FB_DL_SignalDebounce 的边界 —— 去抖是「延迟跳变并对两侧同宽」，本件是
              「短于宽度的整段丢弃且合格脉宽不失真」，两者判据与后果都不同，不可互相替代。
    开源溯源 : 原创实现（T0-1 变体线）。无外部源码参考，码位、抑制计数策略、双侧确认结构 100% 自有。；本件为 IEC 61131-3 标准语义的道莅防御性实现（原创实现，零外部源码复制）。
    本文件内含 : FUNCTION_BLOCK FB_DL_PulseWidthFilter（单 POU，无配套类型）
    依 赖 : 无 DL_ 内部依赖；Standard.library: TON / R_TRIG / F_TRIG
    红线自检 : R1 ✓ 零全局变量与外部变量 ｜ R2 ✓ 零物理 IO 地址
              R3 ✓ 纯 IEC 61131-3 ｜ R4 ✓ 宽度闸 + 计数饱和闸 + 单拍标志先销后置 + 失能直通
              R5 ✓ 全变量中英双语同行注释 ｜ R6 N/A 本件为纯时序件，无顺序状态机（不引入枚举），
              故 03A7 保留预留并在头注释写明理由；7 项红线中「ENUM + CASE + ELSE」对无状态机件为 N/A
              R7 ✓ TON / R_TRIG / F_TRIG 全部在主体最前部无条件刷新，位于任何 IF 之外
              R8 ✓ 最小宽度、告警代理阈值、计数上限全常量化
    错误码   : 16#0001_045A [信息级] 确认窗小于两倍最小任务周期的代理阈值（2ms），只提示不改参数，bError = FALSE
               16#0001_045B [信息级] 预留禁用（不得挪用；本件信息级只用 1 槽，不加强加码 —— R90）
               16#0001_03A5 [故障级] 最小宽度非法已钳至 1ms 继续，bError = TRUE
               16#0001_03A6 [故障级] 抑制计数饱和，统计已失真需复位，bError = TRUE
               16#0001_03A7 [故障级] 预留禁用（本件无状态机，无非法状态分支，故不占实现）
    码位总账 : 16#0001_045A 用 / 16#0001_045B 预留 ｜ 16#0001_03A5 用 / 16#0001_03A6 用 / 16#0001_03A7 预留
    遗留假设 :
        ① 【代理阈值的口径必须明说】库内没有扫描周期引脚（扫描周期由调用方注入的 tDelta 只在
        FB_DL_SamplingTrigger 里出现，本件按派单引脚表不得新增），故无法真正判「tMinWidth < 2 × 扫描周期」。
        本件以 DL_PWF_WARN_MIN = T#2MS（1ms 任务的极限确认窗）作为代理阈值发 045A，
        该代理不能覆盖更慢的任务（如 10ms 任务），须由调用方在参数整定阶段自行核对 —— 未实测，编译门槛未闭合。
        ② 确认窗依赖 TON 的 PT 语义（IN 断开立即清零 ET），为 IEC 语义推导，未逐平台实测。
    修订历史 :
        2026-11-16  v1.0.0  首版，R21 批次 4 入库
        2026-11-16  v1.0.1  R21 终审修复（轻微）：bReset 的引脚注释承诺「上升沿清抑制计数」，主体却写成
                            电平清零 `IF bReset`。HMI 上按住复位按钮不放是常态，此时抑制计数被持续压零，
                            现场会以为「一个窄脉冲都没发生」，而 bRejected 单拍标志仍在正常翻转。
                            现补 rtReset : R_TRIG 实例（与其余实例同段无条件刷新，满足红线 R4）并改为沿判定；
                            同时把引脚注释里并不存在的「饱和标志」措辞改成实情（饱和只为当拍 eErr 报码）。
*)
FUNCTION_BLOCK FB_DL_PulseWidthFilter
VAR_INPUT
    bEnable         : BOOL := TRUE;      // 使能，FALSE 时输出直通输入（旁路）/ enable, FALSE bypasses the filter and follows the input
    bIn             : BOOL;              // 原始信号 / raw input signal
    tMinWidth       : TIME := T#20MS;    // 允许通过的最小脉冲宽度，≤ 0 时钳 1ms [ms] / minimum pulse width that may pass, clamped to one millisecond [ms]
    bReset          : BOOL;              // 上升沿清抑制计数（饱和只是当拍报码，随段 0 预置自动销）/ rising edge clears the reject count, the saturation notice is single scan and clears itself
END_VAR
VAR_OUTPUT
    bOut            : BOOL;              // 过滤后的输出，合格脉冲宽度不失真 / filtered output, the width of an accepted pulse is preserved
    uRejectCount    : UDINT;             // 被吞掉的窄脉冲数 [次] / number of suppressed narrow pulses [count]
    bRejected       : BOOL;              // 本拍是否发生抑制（单拍，恒只活一个扫描周期）/ TRUE on the scan a pulse was suppressed, single scan only
    eErr            : UDINT;             // 错误码，0=正常；16#0001_04XX 信息级 / 16#0001_03XX 故障级 / error id, 0=ok
    bError          : BOOL;              // 故障级标志 / fault flag
END_VAR
VAR
    fbOnDelay       : TON;               // 上升沿确认窗，主体最前部无条件刷新 / high level confirmation timer, refreshed unconditionally at the top
    fbOffDelay      : TON;               // 下降沿确认窗，主体最前部无条件刷新 / low level confirmation timer, refreshed unconditionally at the top
    rtIn            : R_TRIG;            // 输入上升沿，主体最前部无条件刷新 / input rising edge, refreshed unconditionally at the top
    ftIn            : F_TRIG;            // 输入下降沿，主体最前部无条件刷新 / input falling edge, refreshed unconditionally at the top
    rtReset         : R_TRIG;            // 复位上升沿，主体最前部无条件刷新 / reset rising edge, refreshed unconditionally at the top
    bInRaw          : BOOL;              // 使能掩蔽后的输入 / input masked by the enable
    tMinEff         : TIME;              // 钳位后的最小宽度 [ms] / clamped minimum width [ms]
END_VAR
VAR CONSTANT
    DL_PWF_MIN          : TIME := T#1MS;                 // 最小宽度下限 [ms] / minimum width lower bound [ms]
    DL_PWF_WARN_MIN     : TIME := T#2MS;                 // 代理告警阈值（1ms 任务的极限确认窗）[ms] / proxy warning threshold [ms]
    DL_TIME_ZERO        : TIME := T#0S;                  // 零时长哨兵 [ms] / zero duration sentinel [ms]
    DL_UDINT_MAX        : UDINT := 16#FFFF_FFFF;         // 抑制计数上限 [次] / reject count upper bound [count]
    DL_ERR_NONE         : UDINT := 16#0000_0000;         // 无故障 / no error
END_VAR

// 段 0｜错误状态预置与单拍标志清销 / segment 0, preset the error state and clear the single scan flag
eErr      := DL_ERR_NONE;                 // 预置无错误 / preset no error
bError    := FALSE;                       // 预置无故障 / preset no fault
bRejected := FALSE;                       // 单拍标志每拍先销，防「只置不销」/ the single scan flag is cleared first

// 段 1｜宽度闸：非法钳 1ms 继续，不停机 / segment 1, width gate with clamping
IF tMinWidth <= DL_TIME_ZERO THEN
    tMinEff := DL_PWF_MIN;                // 钳到最小宽度 / clamp to the smallest width
    eErr    := 16#0001_03A5;              // 最小宽度非法已钳位（故障级）/ illegal minimum width clamped, fault level
    bError  := TRUE;                      // 置故障标志 / raise the fault flag
ELSE
    tMinEff := tMinWidth;                 // 正常值 / a healthy value
END_IF

// 段 2｜代理阈值提示：确认窗过小时扫描周期可能吃掉确认过程 / segment 2, proxy hint for a very short confirmation window
IF (tMinEff < DL_PWF_WARN_MIN) AND (eErr = DL_ERR_NONE) THEN
    eErr := 16#0001_045A;                 // 确认窗过小提示（信息级，不置 bError）/ short confirmation window hint, info level
END_IF

// 段 3｜定时器与边沿无条件刷新：两只看守的 IN 都串入 bEnable，失能即同步复位 / segment 3, unconditional refresh
bInRaw := bEnable AND bIn;                                    // 使能掩蔽 / mask by the enable
fbOnDelay ( IN := bInRaw,                PT := tMinEff );      // 高电平确认窗 / high level confirmation
fbOffDelay( IN := (NOT bInRaw) AND bEnable, PT := tMinEff );   // 低电平确认窗，失能时同步复位 / low level confirmation, reset while disabled
rtIn      ( CLK := bInRaw );                                   // 输入上升沿 / input rising edge
ftIn      ( CLK := bInRaw );                                   // 输入下降沿 / input falling edge
rtReset   ( CLK := bReset );                                   // 复位上升沿，与其余实例同段无条件刷新 / reset rising edge, refreshed unconditionally in the same segment

// 段 4｜复位沿：清抑制统计（引脚注释承诺「上升沿」，故必须真做沿判定，禁用电平清零）/ segment 4, the reset edge clears the suppression statistics
IF rtReset.Q THEN
    uRejectCount := 0;                    // 计数清零 / clear the count
END_IF

// 段 5｜失能直通：旁路时不得留门控残影 / segment 5, bypass without any residual gating
IF NOT bEnable THEN
    bOut := bIn;                          // 直通输入 / follow the input directly
ELSE
    // 段 6｜双侧确认搬运：高电平确认满才置高，低电平确认满才置低，故输出宽度与输入同宽 / segment 6, two sided transfer
    IF fbOnDelay.Q THEN
        bOut := TRUE;                     // 高电平已维持满最小宽度 / the high level lasted long enough
    END_IF
    IF fbOffDelay.Q THEN
        bOut := FALSE;                    // 低电平已维持满最小宽度 / the low level lasted long enough
    END_IF

    // 段 7｜窄脉冲判定：高电平未确认即回落 → 窄高脉冲；低电平未确认即回升 → 窄低脉冲 / segment 7, narrow pulse detection
    IF ftIn.Q AND (NOT bOut) THEN
        bRejected := TRUE;                // 窄高脉冲：上升后未确认就掉了 / a narrow high pulse fell before confirmation
    END_IF
    IF rtIn.Q AND bOut THEN
        bRejected := TRUE;                // 窄低脉冲：下降后未确认就回来了 / a narrow low pulse rose before confirmation
    END_IF

    // 段 8｜抑制计数：饱和后不再递增并报故障（统计已失真需复位）/ segment 8, reject counting with saturation
    IF bRejected THEN
        IF uRejectCount >= DL_UDINT_MAX THEN
            eErr   := 16#0001_03A6;       // 抑制计数饱和（故障级）/ reject count saturated, fault level
            bError := TRUE;               // 置故障标志 / raise the fault flag
        ELSE
            uRejectCount := uRejectCount + 1;   // 计数递增 / increment the count
        END_IF
    END_IF
END_IF
END_FUNCTION_BLOCK
